(* Logix 5000 project; controller NWGG 1756-L72 rev 35.12; software revision 35.00; part 13 of 19 *)
(* tags used below, declared in another part *)
   tmrWeightTest : TIMER;
   Weight_Seed : DINT;
   _103_TANK_42_RECEIVING_LEG_RUNNING : BOOL;
   _106_TANK_17_AUGER_RUNNING : BOOL;
   _107_TANKS_1THRU7_SOUTH_RUNNING : BOOL;
   _108_CENTER_BELT_RUNNING : BOOL;
   _109_RAW_RECEIVING_NORTH_BELT_RUNNING : BOOL;
   _110_TANK_16_AUGER_RUNNING : BOOL;
   _113_HIGHROLLER_TANKS_11TO15_RUNNING : BOOL;
   _114_TANKS_1THRU7_NORTH_RUNNING : BOOL;
   _11_TANK_41_42_HIGHROLLER_RUNNING : BOOL;
   _123_CLEAN_LEG_RUNNING : BOOL;
   _1_CLEAN_SEED_UPPER_BELT_RUNNING : BOOL;
   _35_JUMP_LEG_RUNNING : BOOL;
   _3_LOWER_TANK_CONVAYOR_24TO26_RUNNING : BOOL;
   _43_SCREENINGS_LEG_RUNNING : BOOL;
   _4_LOWER_TANK_CONVAYOR_21TO23_RUNNING : BOOL;
   _5_LOWER_CROSS_BELT_RUNNING : BOOL;
   _701_TRUCK_REVERSING_BELT_RUNNING : BOOL;
   _703_TREATER_JUMP_BELT_RUNNING : BOOL;
   _9_TREATER_CONVAYOR_RUNNING : BOOL;
   Analog : AI[160];
   Calibration_Max : REAL;
   InEUMax : REAL;
   TestTag : REAL;
   Truck_Scales : udt_Truck_Scale[2];
(* MainProgram, continued *)

ROUTINE Totals   (* function block diagram *)
   SHEET 1
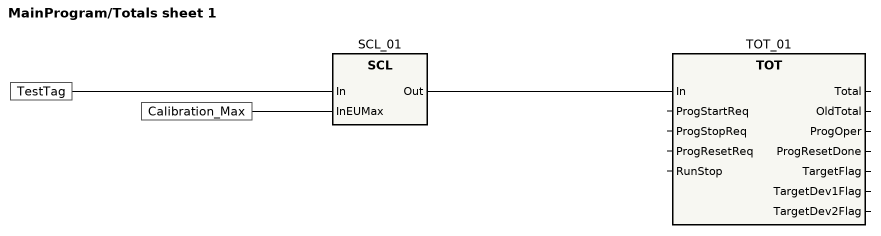
   SCL_01 : SCL(In := TestTag, InEUMax := Calibration_Max);
   TOT_01 : TOT(In := SCL_01.Out);   // unwired pins: ProgStartReq ProgStopReq ProgResetReq Total OldTotal ProgOper RunStop ProgResetDone TargetFlag TargetDev1Flag TargetDev2Flag
END_ROUTINE

ROUTINE VERIFACATION   (* ladder *)
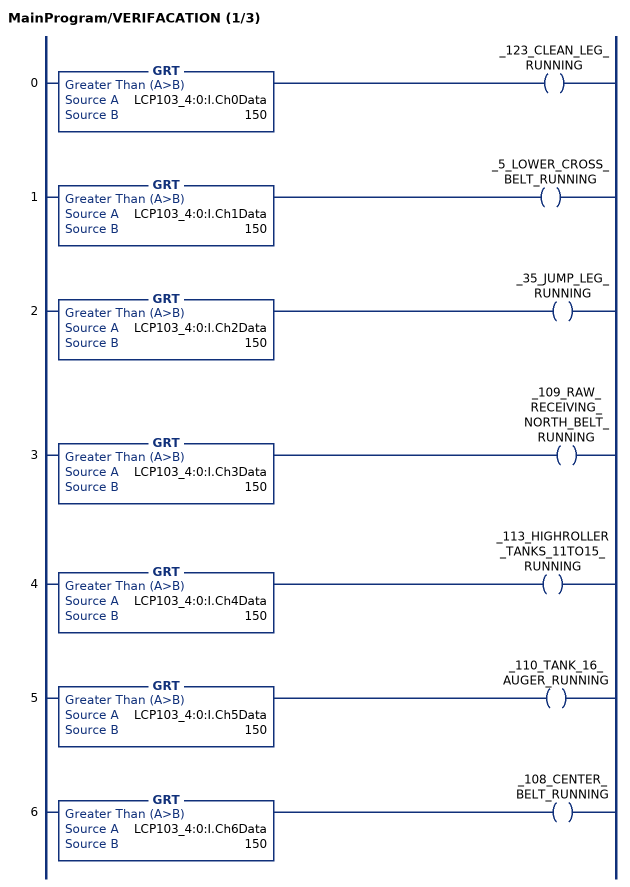
   0: GRT(LCP103_4:0:I.Ch0Data,150)OTE(_123_CLEAN_LEG_RUNNING);
   1: GRT(LCP103_4:0:I.Ch1Data,150)OTE(_5_LOWER_CROSS_BELT_RUNNING);
   2: GRT(LCP103_4:0:I.Ch2Data,150)OTE(_35_JUMP_LEG_RUNNING);
   3: GRT(LCP103_4:0:I.Ch3Data,150)OTE(_109_RAW_RECEIVING_NORTH_BELT_RUNNING);
   4: GRT(LCP103_4:0:I.Ch4Data,150)OTE(_113_HIGHROLLER_TANKS_11TO15_RUNNING);
   5: GRT(LCP103_4:0:I.Ch5Data,150)OTE(_110_TANK_16_AUGER_RUNNING);
   6: GRT(LCP103_4:0:I.Ch6Data,150)OTE(_108_CENTER_BELT_RUNNING);
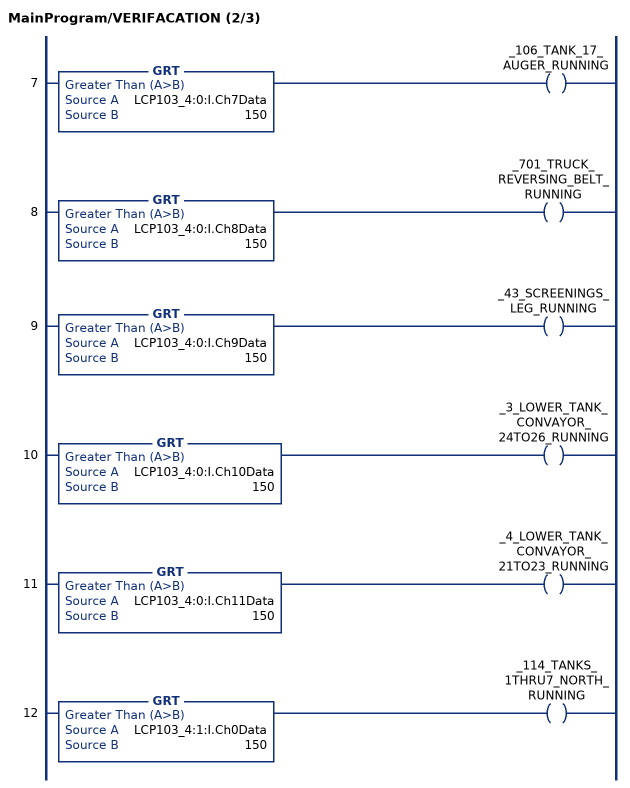
   7: GRT(LCP103_4:0:I.Ch7Data,150)OTE(_106_TANK_17_AUGER_RUNNING);
   8: GRT(LCP103_4:0:I.Ch8Data,150)OTE(_701_TRUCK_REVERSING_BELT_RUNNING);
   9: GRT(LCP103_4:0:I.Ch9Data,150)OTE(_43_SCREENINGS_LEG_RUNNING);
   10: GRT(LCP103_4:0:I.Ch10Data,150)OTE(_3_LOWER_TANK_CONVAYOR_24TO26_RUNNING);
   11: GRT(LCP103_4:0:I.Ch11Data,150)OTE(_4_LOWER_TANK_CONVAYOR_21TO23_RUNNING);
   12: GRT(LCP103_4:1:I.Ch0Data,150)OTE(_114_TANKS_1THRU7_NORTH_RUNNING);
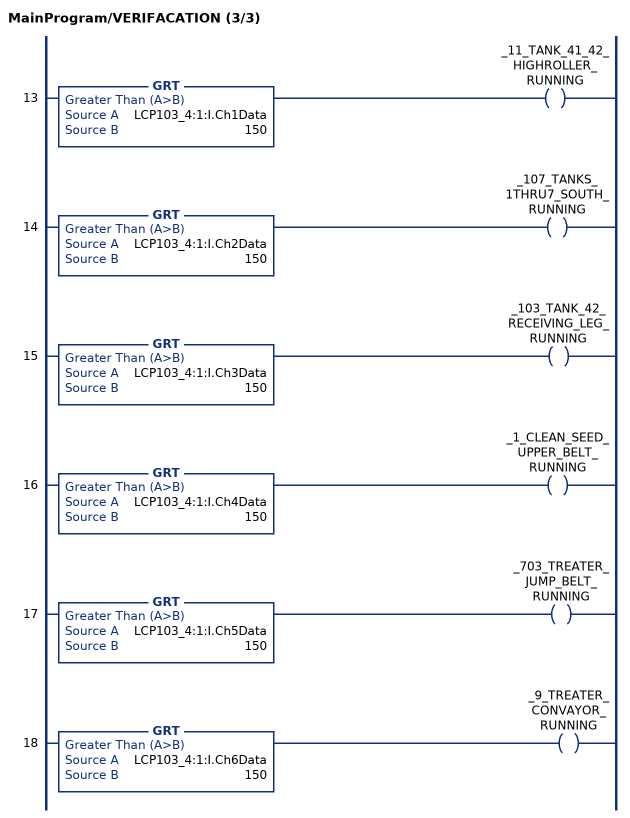
   13: GRT(LCP103_4:1:I.Ch1Data,150)OTE(_11_TANK_41_42_HIGHROLLER_RUNNING);
   14: GRT(LCP103_4:1:I.Ch2Data,150)OTE(_107_TANKS_1THRU7_SOUTH_RUNNING);
   15: GRT(LCP103_4:1:I.Ch3Data,150)OTE(_103_TANK_42_RECEIVING_LEG_RUNNING);
   16: GRT(LCP103_4:1:I.Ch4Data,150)OTE(_1_CLEAN_SEED_UPPER_BELT_RUNNING);
   17: GRT(LCP103_4:1:I.Ch5Data,150)OTE(_703_TREATER_JUMP_BELT_RUNNING);
   18: GRT(LCP103_4:1:I.Ch6Data,150)OTE(_9_TREATER_CONVAYOR_RUNNING);
END_ROUTINE

ROUTINE Weigh_Scales   (* ladder *)
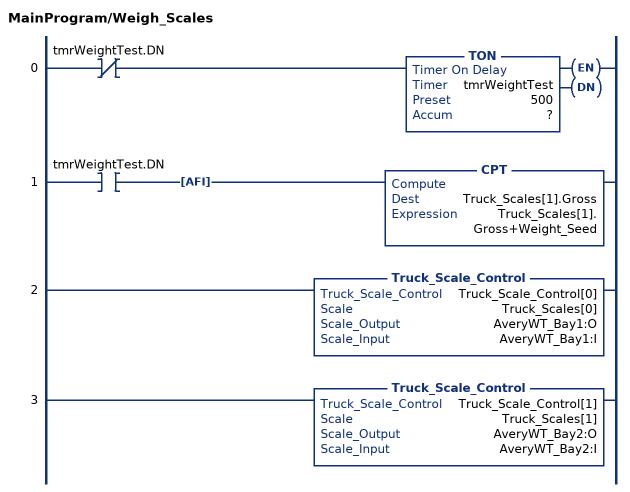
   0: XIO(tmrWeightTest.DN)TON(tmrWeightTest,?,?);
   1: XIC(tmrWeightTest.DN)AFI()CPT(Truck_Scales[1].Gross,Truck_Scales[1].Gross+Weight_Seed);
   2: Truck_Scale_Control(Truck_Scale_Control[0],Truck_Scales[0],AveryWT_Bay1:O,AveryWT_Bay1:I);
   3: Truck_Scale_Control(Truck_Scale_Control[1],Truck_Scales[1],AveryWT_Bay2:O,AveryWT_Bay2:I);
END_ROUTINE
END_PROGRAM

PROGRAM Scale   (* main routine MainRoutine *)
VAR
   ctlAddTime : CONTROL[2];
   ctrWtArray : COUNTER[2] := ([0].DN := 1, [1].DN := 1);
   Cur_Weight : REAL[2];
   Cur_Weight_Array_Idx : DINT := 16;
   Current_Gross : DINT[2];
   Current_Weight : REAL;
   Prev_Weight : REAL[2];
   Scale_Rate : REAL[2];
   Scale_Test_Rate_Mlt : DINT;
   ScaleIDX : DINT := 2;
   ShiftIDX : DINT := 20;
   TestRate : REAL[2];
   Time_Array : DINT[2,10] := ([0,0] := 9, [0,1] := 9, [0,2] := 10, [0,3] := 10, [0,4] := 8, [0,5] := 10, [0,6] := 9, [0,7] := 9, [0,8] := 9, [1,0] := 10, [1,1] := 9, [1,2] := 10, [1,3] := 10, [1,4] := 9, [1,5] := 10, [1,6] := 8, [1,7] := 10, [1,8] := 9);
   tmrRate : TIMER[2] := ([0].PRE := 1000, [0].ACC := 109, [0].EN := 1, [0].TT := 1, [1].PRE := 1000, [1].ACC := 126, [1].EN := 1, [1].TT := 1);
   tmrTestRate : TIMER[2] := ([1].ACC := 15, [1].EN := 1, [1].DN := 1);
   Total_Time : DINT[2];
   Weight_Array : REAL[2,40];
   Weight_Array_Idx : DINT[2] := ([0] := 14, [1] := 17);
   Weight_Array_Max : REAL[2];
   Weight_Sum : REAL[2];
END_VAR

ROUTINE AddWeights   (* ladder *)
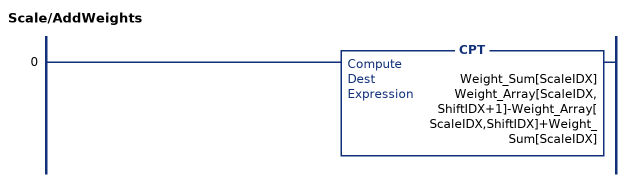
   0: CPT(Weight_Sum[ScaleIDX],Weight_Array[ScaleIDX,ShiftIDX+1]-Weight_Array[ScaleIDX,ShiftIDX]+Weight_Sum[ScaleIDX]);
END_ROUTINE

ROUTINE MainRoutine   (* ladder *)
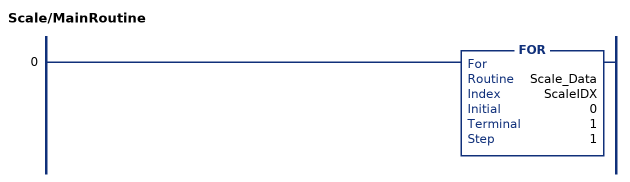
   0: FOR(Scale_Data,ScaleIDX,0,1,1);
END_ROUTINE

ROUTINE Scale_Data   (* ladder *)
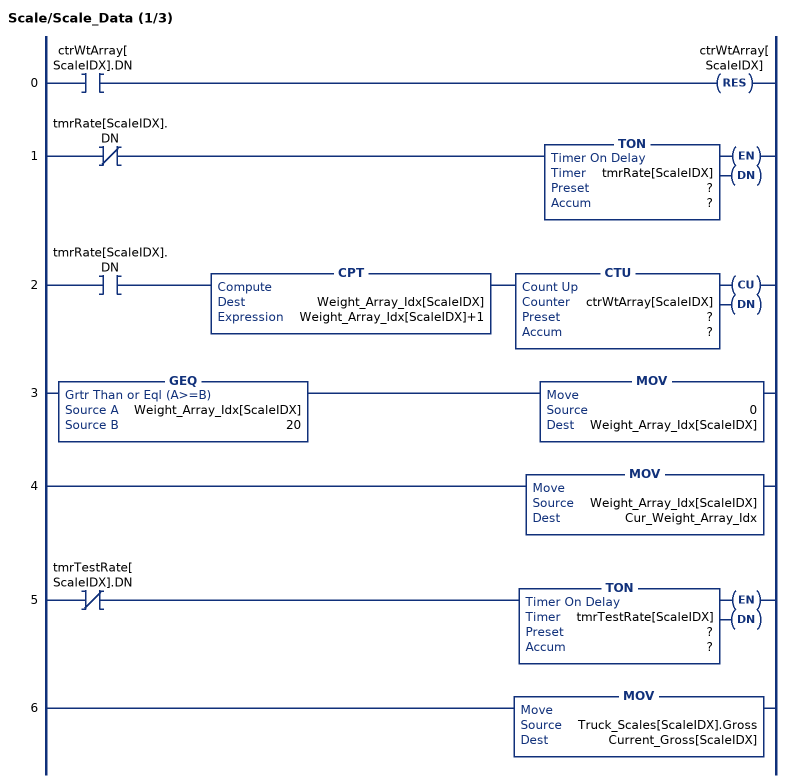
   0: XIC(ctrWtArray[ScaleIDX].DN)RES(ctrWtArray[ScaleIDX]);
   1: XIO(tmrRate[ScaleIDX].DN)TON(tmrRate[ScaleIDX],?,?);
   2: XIC(tmrRate[ScaleIDX].DN)CPT(Weight_Array_Idx[ScaleIDX],Weight_Array_Idx[ScaleIDX]+1)CTU(ctrWtArray[ScaleIDX],?,?);
   3: GEQ(Weight_Array_Idx[ScaleIDX],20)MOV(0,Weight_Array_Idx[ScaleIDX]);
   4: MOV(Weight_Array_Idx[ScaleIDX],Cur_Weight_Array_Idx);
   5: XIO(tmrTestRate[ScaleIDX].DN)TON(tmrTestRate[ScaleIDX],?,?);
   6: MOV(Truck_Scales[ScaleIDX].Gross,Current_Gross[ScaleIDX]);
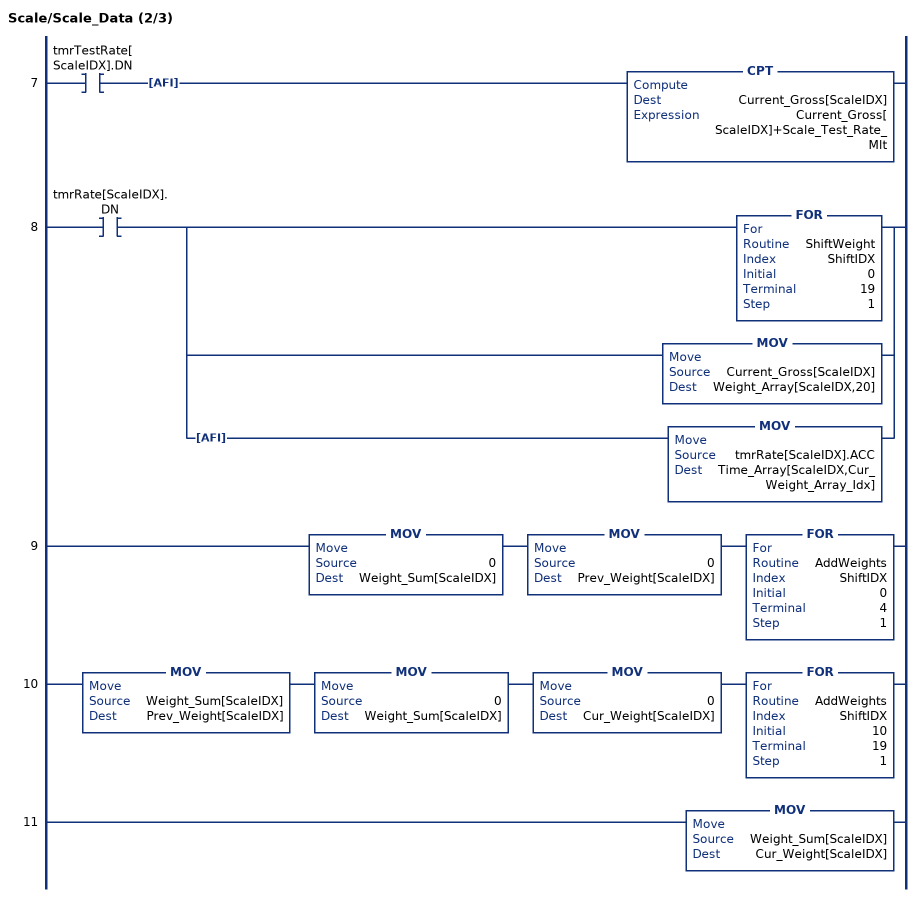
   7: XIC(tmrTestRate[ScaleIDX].DN)AFI()CPT(Current_Gross[ScaleIDX],Current_Gross[ScaleIDX]+Scale_Test_Rate_Mlt);
   8: XIC(tmrRate[ScaleIDX].DN)[FOR(ShiftWeight,ShiftIDX,0,19,1) ,MOV(Current_Gross[ScaleIDX],Weight_Array[ScaleIDX,20]) ,AFI() MOV(tmrRate[ScaleIDX].ACC,Time_Array[ScaleIDX,Cur_Weight_Array_Idx]) ];
   9: MOV(0,Weight_Sum[ScaleIDX])MOV(0,Prev_Weight[ScaleIDX])FOR(AddWeights,ShiftIDX,0,4,1);
   10: MOV(Weight_Sum[ScaleIDX],Prev_Weight[ScaleIDX])MOV(0,Weight_Sum[ScaleIDX])MOV(0,Cur_Weight[ScaleIDX])FOR(AddWeights,ShiftIDX,10,19,1);
   11: MOV(Weight_Sum[ScaleIDX],Cur_Weight[ScaleIDX]);
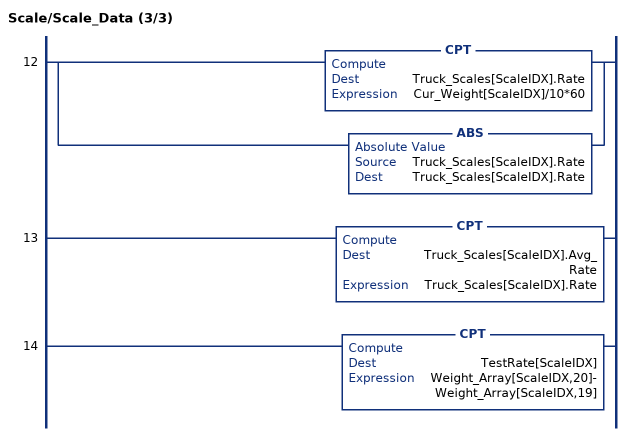
   12: [CPT(Truck_Scales[ScaleIDX].Rate,Cur_Weight[ScaleIDX]/10*60) ,ABS(Truck_Scales[ScaleIDX].Rate,Truck_Scales[ScaleIDX].Rate) ];
   13: CPT(Truck_Scales[ScaleIDX].Avg_Rate,Truck_Scales[ScaleIDX].Rate);
   14: CPT(TestRate[ScaleIDX],Weight_Array[ScaleIDX,20]-Weight_Array[ScaleIDX,19]);
END_ROUTINE

ROUTINE ShiftWeight   (* ladder *)
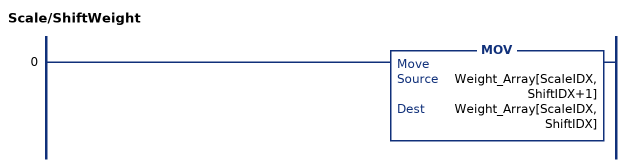
   0: MOV(Weight_Array[ScaleIDX,ShiftIDX+1],Weight_Array[ScaleIDX,ShiftIDX]);
END_ROUTINE
END_PROGRAM

PROGRAM SeedLoadoutMain   (* main routine MainRoutine *)
VAR
   Accept_Bin_Cal : BOOL;
   Air_Gates_Opened : BOOL;
   All_Stop : BOOL;
   ALM_Air_Gate_Failed_Open_Bin0 : ALARM_DIGITAL;
   ALM_Air_Gate_Failed_Open_Bin1 : ALARM_DIGITAL;
   ALM_Air_Gate_Failed_Open_Bin10 : ALARM_DIGITAL;
   ALM_Air_Gate_Failed_Open_Bin11 : ALARM_DIGITAL;
   ALM_Air_Gate_Failed_Open_Bin12 : ALARM_DIGITAL;
   ALM_Air_Gate_Failed_Open_Bin13 : ALARM_DIGITAL;
   ALM_Air_Gate_Failed_Open_Bin14 : ALARM_DIGITAL;
   ALM_Air_Gate_Failed_Open_Bin15 : ALARM_DIGITAL;
   ALM_Air_Gate_Failed_Open_Bin16 : ALARM_DIGITAL;
   ALM_Air_Gate_Failed_Open_Bin17 : ALARM_DIGITAL;
   ALM_Air_Gate_Failed_Open_Bin18 : ALARM_DIGITAL;
   ALM_Air_Gate_Failed_Open_Bin19 : ALARM_DIGITAL;
   ALM_Air_Gate_Failed_Open_Bin2 : ALARM_DIGITAL;
   ALM_Air_Gate_Failed_Open_Bin20 : ALARM_DIGITAL;
   ALM_Air_Gate_Failed_Open_Bin21 : ALARM_DIGITAL;
   ALM_Air_Gate_Failed_Open_Bin22 : ALARM_DIGITAL;
   ALM_Air_Gate_Failed_Open_Bin23 : ALARM_DIGITAL;
   ALM_Air_Gate_Failed_Open_Bin24 : ALARM_DIGITAL;
   ALM_Air_Gate_Failed_Open_Bin25 : ALARM_DIGITAL;
   ALM_Air_Gate_Failed_Open_Bin26 : ALARM_DIGITAL;
   ALM_Air_Gate_Failed_Open_Bin27 : ALARM_DIGITAL;
   ALM_Air_Gate_Failed_Open_Bin28 : ALARM_DIGITAL;
   ALM_Air_Gate_Failed_Open_Bin3 : ALARM_DIGITAL;
   ALM_Air_Gate_Failed_Open_Bin4 : ALARM_DIGITAL;
   ALM_Air_Gate_Failed_Open_Bin5 : ALARM_DIGITAL;
   ALM_Air_Gate_Failed_Open_Bin6 : ALARM_DIGITAL;
   ALM_Air_Gate_Failed_Open_Bin7 : ALARM_DIGITAL;
   ALM_Air_Gate_Failed_Open_Bin8 : ALARM_DIGITAL;
   ALM_Air_Gate_Failed_Open_Bin9 : ALARM_DIGITAL;
   ALM_K_Valve1_Treat_Failed : ALARM_DIGITAL;
   ALM_KValve0_Clean_Failed : ALARM_DIGITAL;
   ALM_KValve0_Treat_Failed : ALARM_DIGITAL;
   ALM_KValve1_Clean_Failed : ALARM_DIGITAL;
   ALM_NOT_USED : ALARM_DIGITAL;
   ALM_OVRAMP_Belt10 : ALARM_DIGITAL;
   ALM_OVRAMP_Belt11 : ALARM_DIGITAL;
   ALM_OVRAMP_Belt2 : ALARM_DIGITAL;
   ALM_OVRAMP_Belt3 : ALARM_DIGITAL;
   ALM_OVRAMP_Belt4 : ALARM_DIGITAL;
   ALM_OVRAMP_Belt5 : ALARM_DIGITAL;
   ALM_OVRAMP_Belt6 : ALARM_DIGITAL;
   ALM_OVRAMP_Belt7 : ALARM_DIGITAL;
   ALM_OVRAMP_Belt8 : ALARM_DIGITAL;
   ALM_OVRAMP_Belt9 : ALARM_DIGITAL;
   ALM_OVRAMP_CPLeg : ALARM_DIGITAL;
   ALM_PLUG_Belt1 : ALARM_DIGITAL;
   ALM_PLUG_Belt10 : ALARM_DIGITAL;
   ALM_PLUG_Belt11 : ALARM_DIGITAL;
   ALM_PLUG_Belt2 : ALARM_DIGITAL;
   ALM_PLUG_Belt3 : ALARM_DIGITAL;
   ALM_PLUG_Belt4 : ALARM_DIGITAL;
   ALM_PLUG_Belt5 : ALARM_DIGITAL;
   ALM_PLUG_Belt6 : ALARM_DIGITAL;
   ALM_PLUG_Belt7 : ALARM_DIGITAL;
   ALM_PLUG_Belt8 : ALARM_DIGITAL;
   ALM_PLUG_Belt9 : ALARM_DIGITAL;
   ALM_PLUG_CPLeg : ALARM_DIGITAL;
   ALM_SLP10_Belt1 : ALARM_DIGITAL;
   ALM_SLP10_Belt10 : ALARM_DIGITAL;
   ALM_SLP10_Belt11 : ALARM_DIGITAL;
   ALM_SLP10_Belt2 : ALARM_DIGITAL;
   ALM_SLP10_Belt3 : ALARM_DIGITAL;
   ALM_SLP10_Belt4 : ALARM_DIGITAL;
   ALM_SLP10_Belt5 : ALARM_DIGITAL;
   ALM_SLP10_Belt6 : ALARM_DIGITAL;
   ALM_SLP10_Belt7 : ALARM_DIGITAL;
   ALM_SLP10_Belt8 : ALARM_DIGITAL;
   ALM_SLP10_Belt9 : ALARM_DIGITAL;
   ALM_SLP10_CPLeg : ALARM_DIGITAL;
   ALM_SLP20_Belt1 : ALARM_DIGITAL;
   ALM_SLP20_Belt10 : ALARM_DIGITAL;
   ALM_SLP20_Belt11 : ALARM_DIGITAL;
   ALM_SLP20_Belt2 : ALARM_DIGITAL;
   ALM_SLP20_Belt3 : ALARM_DIGITAL;
   ALM_SLP20_Belt4 : ALARM_DIGITAL;
   ALM_SLP20_Belt5 : ALARM_DIGITAL;
   ALM_SLP20_Belt6 : ALARM_DIGITAL;
   ALM_SLP20_Belt7 : ALARM_DIGITAL;
   ALM_SLP20_Belt8 : ALARM_DIGITAL;
   ALM_SLP20_Belt9 : ALARM_DIGITAL;
   ALM_SLP20_CPLeg : ALARM_DIGITAL;
   ALM_WONT_START_Belt1 : ALARM_DIGITAL;
   ALM_WONT_START_Belt10 : ALARM_DIGITAL;
   ALM_WONT_START_Belt11 : ALARM_DIGITAL;
   ALM_WONT_START_Belt2 : ALARM_DIGITAL;
   ALM_WONT_START_Belt3 : ALARM_DIGITAL;
   ALM_WONT_START_Belt4 : ALARM_DIGITAL;
   ALM_WONT_START_Belt5 : ALARM_DIGITAL;
   ALM_WONT_START_Belt6 : ALARM_DIGITAL;
   ALM_WONT_START_Belt7 : ALARM_DIGITAL;
   ALM_WONT_START_Belt8 : ALARM_DIGITAL;
   ALM_WONT_START_Belt9 : ALARM_DIGITAL;
   ALM_WONT_START_CPLeg : ALARM_DIGITAL;
   Always_Off : BOOL;
   Andco_Auto_Mode : BOOL;
   Andco_Rate : DINT;
   Auto_Mode : BOOL := 1;
   Auto_Mode_ONS : BOOL;
   Auto_Start_Reversing_Belt_Fans : BOOL;
   Auto_Start_Treatment : BOOL;
   Auto_Stop_Clean : BOOL;
   Auto_Stop_Clean_Belt_11 : BOOL;
   Auto_Stop_Transfer : BOOL;
   Auto_Stop_Treat : BOOL;
   Available_For_Clean_Loadout : DINT := 536870911;
   Available_For_Treat_Loadout : DINT := 536870911;
   b3 : ALARM_DIGITAL;
   B_Offset : REAL;
   Batch_Status : DINT;
   BC_3_Belt_Required : BOOL;
   BC_9_Interlock : BOOL;
   Belt : udt_Motor[16] := ([0].Motor_Start.Auto_Stop_Delay := 5000, [1].Motor_Start.Auto_Stop_Delay := 5000, [1].Motor_Control.Spd_10_Pct := 1, [1].Motor_Control.Motor_Amps := -0.32500002, [1].Motor_Control.Motor_Batch_Ready := 1, [1].Motor_Control.Motor_Batch_Ready_Clean := 1, [1].Motor_Control.Motor_Batch_Ready_Treat := 1, [1].Motor_Control.Motor_Batch_Ready_Transfer := 1, [1].Motor_Config.Definition := 'Middle Concrete', [1].Motor_Config.Wind_Up_Time := 3000, [1].Motor_Config.Stop_At_SLP20 := 1, [1].Motor_Config.Stop_At_Max_Amps := 1, [1].Motor_Config.Max_Amps := 1000.0, [2].Motor_Start.Auto_Stop_Delay := 5000, [2].Motor_Control.Spd_10_Pct := 1, [2].Motor_Control.Motor_Amps := -0.4125, [2].Motor_Control.Motor_Batch_Ready := 1, [2].Motor_Control.Motor_Batch_Ready_Clean := 1, [2].Motor_Control.Motor_Batch_Ready_Treat := 1, [2].Motor_Control.Motor_Batch_Ready_Transfer := 1, [2].Motor_Config.Definition := 'North Concrete', [2].Motor_Config.Wind_Up_Time := 3000, [2].Motor_Config.Stop_At_SLP20 := 1, [3].Motor_Start.Auto_Stop_Delay := 5000, [3].Motor_Control.Spd_10_Pct := 1, [3].Motor_Control.Motor_Amps := -0.5125, [3].Motor_Control.Motor_Batch_Ready := 1, [3].Motor_Control.Motor_Batch_Ready_Clean := 1, [3].Motor_Control.Motor_Batch_Ready_Treat := 1, [3].Motor_Control.Motor_Batch_Ready_Transfer := 1, [3].Motor_Config.Definition := 'South Concrete', [3].Motor_Config.Wind_Up_Time := 3000, [3].Motor_Config.Stop_At_SLP20 := 1, [4].Motor_Start.Auto_Stop_Delay := 5000, [4].Motor_Control.Motor_Amps := -0.05285539, [4].Motor_Control.Motor_Batch_Ready := 1, [4].Motor_Control.Motor_Batch_Ready_Clean := 1, [4].Motor_Control.Motor_Batch_Ready_Treat := 1, [4].Motor_Control.Motor_Batch_Ready_Transfer := 1, [4].Motor_Config.Definition := 'Reversing', [4].Motor_Config.Wind_Up_Time := 6000, [4].Motor_Config.Stop_At_SLP20 := 1, [5].Motor_Start.Auto_Stop_Delay := 5000, [5].Motor_Control.Spd_10_Pct := 1, [5].Motor_Control.Motor_Amps := 0.018231237, [5].Motor_Control.Motor_Batch_Ready := 1, [5].Motor_Control.Motor_Batch_Ready_Clean := 1, [5].Motor_Control.Motor_Batch_Ready_Treat := 1, [5].Motor_Control.Motor_Batch_Ready_Transfer := 1, [5].Motor_Config.Definition := 'Treat Jump', [5].Motor_Config.Wind_Up_Time := 3000, [5].Motor_Config.Stop_At_SLP20 := 1, [6].Motor_Start.Auto_Stop_Delay := 5000, [6].Motor_Control.Spd_10_Pct := 1, [6].Motor_Control.Motor_Amps := 0.013243717, [6].Motor_Control.Motor_Batch_Ready := 1, [6].Motor_Control.Motor_Batch_Ready_Clean := 1, [6].Motor_Control.Motor_Batch_Ready_Treat := 1, [6].Motor_Control.Motor_Batch_Ready_Transfer := 1, [6].Motor_Config.Definition := 'Clean Jump',
        [6].Motor_Config.Wind_Up_Time := 3000, [6].Motor_Config.Stop_At_SLP20 := 1, [6].Motor_Config.Plugged_Sensor_Disabled := 1, [7].Motor_Start.Auto_Stop_Delay := 5000, [7].Motor_Control.Spd_10_Pct := 1, [7].Motor_Control.Motor_Amps := -0.23403546, [7].Motor_Control.Motor_Batch_Ready := 1, [7].Motor_Control.Motor_Batch_Ready_Clean := 1, [7].Motor_Control.Motor_Batch_Ready_Treat := 1, [7].Motor_Control.Motor_Batch_Ready_Transfer := 1, [7].Motor_Config.Definition := 'BC-9', [7].Motor_Config.Wind_Up_Time := 3000, [7].Motor_Config.Stop_At_SLP20 := 1, [7].Motor_Config.Plugged_Sensor_Disabled := 1, [8].Motor_Start.Auto_Stop_Delay := 5000, [8].Motor_Control.Spd_20_Pct := 1, [8].Motor_Control.Motor_Amps := 0.001667556, [8].Motor_Control.Motor_Batch_Ready := 1, [8].Motor_Control.Motor_Batch_Ready_Clean := 1, [8].Motor_Control.Motor_Batch_Ready_Treat := 1, [8].Motor_Control.Motor_Batch_Ready_Transfer := 1, [8].Motor_Config.Definition := 'BC-4', [8].Motor_Config.Wind_Up_Time := 3000, [8].Motor_Config.Speed_Sensor_Disabled := 1, [8].Motor_Config.Plugged_Sensor_Disabled := 1, [9].Motor_Start.Auto_Stop_Delay := 5000, [9].Motor_Control.Spd_20_Pct := 1, [9].Motor_Control.Motor_Amps := 0.033333335, [9].Motor_Control.Motor_Batch_Ready := 1, [9].Motor_Control.Motor_Batch_Ready_Clean := 1, [9].Motor_Control.Motor_Batch_Ready_Treat := 1, [9].Motor_Control.Motor_Batch_Ready_Transfer := 1, [9].Motor_Config.Definition := 'BC-3', [9].Motor_Config.Wind_Up_Time := 3000, [10].Motor_Start.Auto_Stop_Delay := 5000, [10].Motor_Control.Spd_20_Pct := 1, [10].Motor_Control.Motor_Amps := 0.016583197, [10].Motor_Control.Motor_Batch_Ready := 1, [10].Motor_Control.Motor_Batch_Ready_Clean := 1, [10].Motor_Control.Motor_Batch_Ready_Treat := 1, [10].Motor_Control.Motor_Batch_Ready_Transfer := 1, [10].Motor_Config.Definition := 'High Roller', [10].Motor_Config.Wind_Up_Time := 3000, [11].Motor_Start.Auto_Stop_Delay := 5000, [11].Motor_Control.Spd_20_Pct := 1, [11].Motor_Control.Motor_Amps := -0.008290774, [11].Motor_Control.Motor_Batch_Ready := 1, [11].Motor_Control.Motor_Batch_Ready_Clean := 1, [11].Motor_Control.Motor_Batch_Ready_Treat := 1, [11].Motor_Control.Motor_Batch_Ready_Transfer := 1, [11].Motor_Config.Definition := 'BC-5', [11].Motor_Config.Wind_Up_Time := 3000, [12].Motor_Start.Auto_Stop_Delay := 5000);
   Belt_Amps_Scale : SCALE[11];
   Belt_Gate_Leg_ON : BOOL;
   Belts_Ready : BOOL := 1;
   Belts_Running : BOOL;
   Bin_Cal : BOOL;
   Bin_Cal_IDX : DINT := -1;
   Bin_Calibration : BOOL;
   Bin_Clean_Pause : BOOL;
   Bin_Gate_Test : BOOL := 1;
   Bin_Loadout_Control : Loadout_Bin_Control[29] := ([0].Use_Bindicator := 1, [0].RawAnalogTag := 10270, [1].RawAnalogTag := 9993, [2].Use_Bindicator := 1, [2].RawAnalogTag := 8109, [3].RawAnalogTag := 3610, [4].RawAnalogTag := 7694, [5].RawAnalogTag := 5041, [6].RawAnalogTag := 9661, [7].RawAnalogTag := 9884, [8].RawAnalogTag := 10717, [9].RawAnalogTag := 9078, [10].RawAnalogTag := 8853, [11].RawAnalogTag := 9587, [12].RawAnalogTag := 7657, [13].RawAnalogTag := 9087, [14].RawAnalogTag := 9078, [15].RawAnalogTag := 8853, [16].Use_Bindicator := 1, [16].RawAnalogTag := 14748, [17].Use_Bindicator := 1, [17].RawAnalogTag := 15440, [18].Use_Bindicator := 1, [18].RawAnalogTag := 14244, [19].Use_Bindicator := 1, [19].RawAnalogTag := 13454, [20].Use_Bindicator := 1, [20].RawAnalogTag := 14460, [21].Use_Auger_Relay := 1, [21].Use_Bindicator := 1, [21].RawAnalogTag := 6343, [22].Use_Auger_Relay := 1, [22].Use_Bindicator := 1, [22].RawAnalogTag := 8758, [23].Use_Bindicator := 1, [23].RawAnalogTag := 15944, [24].Use_Bindicator := 1, [24].RawAnalogTag := 15184, [25].Use_Bindicator := 1, [25].RawAnalogTag := 15745, [26].Use_Bindicator := 1, [26].RawAnalogTag := 15279, [27].Use_Bindicator := 1, [27].RawAnalogTag := 14611, [28].Use_Bindicator := 1, [28].RawAnalogTag := 15145);
   Bin_Open_test : BOOL := 1;
   Bin_Transfer_Pause : BOOL;
   Bin_Treat_Pause : BOOL;
   Bin_Use_Index : DINT;
   Bin_Variety_Id : STRING[30] := ([0] := '823048', [1] := '823054', [2] := '823058', [3] := '823038', [4] := '823082', [5] := '823090', [6] := '823054', [7] := '823001', [9] := '873002', [10] := '873002', [11] := '873003', [12] := '823072', [16] := '823098', [17] := '843022', [19] := '822087', [20] := '803003', [21] := '823093', [22] := '843036', [23] := '843001', [24] := '843002', [25] := '843022', [26] := '803003', [27] := '823087', [28] := '803021');
   Bins_Rqd : BOOL;
   Blow_Out_Time : DINT;
   Blow_Out_Time_Remaining : REAL := -0.016;
   Blower_707_Running : BOOL;
   boolTransferTime : BOOL;
   Cal_Bin_Status : DINT;
   Cal_Done : BOOL;
   Calibrate_Mode : BOOL;
   Cancel_Bin_Config : BOOL;
   ckIDX : DINT := 29;
   Clean_Batch_Status : DINT;
   Clean_Bin_Gates_Opened : BOOL := 1;
   Clean_Interlock : BOOL;
   Clean_K_Relay_Not_Used : BOOL := 1;
   Clean_Load_Requested : BOOL;
   Clean_Scale_Target : DINT;
   Clean_Scale_Unavailable : BOOL;
   CleanHours : DINT;
   CleanMinuets : DINT;
   CleanSeconds : DINT;
   cntCleanTime : COUNTER := (PRE := 1);
   cntTest : COUNTER := (PRE := 100, ACC := 4);
   cntTransferTime : COUNTER := (PRE := 1);
   cntTreatTime : COUNTER := (PRE := 1);
   Concrete_Belts_Ready : BOOL;
   Concrete_Bin_Timing_Offset : DINT := 5;
   Concrete_Clean_Belts_Ready : BOOL;
   Concrete_Fan_Start : BOOL;
   Concrete_Leg : udt_Motor := (Motor_Start.Auto_Stop_Delay := 1, Motor_Control.Spd_20_Pct := 1, Motor_Control.Spd_10_Pct := 1, Motor_Control.Motor_Amps := -0.4625, Motor_Control.Motor_Batch_Ready_Clean := 1, Motor_Control.Motor_Batch_Ready_Treat := 1, Motor_Control.Motor_Batch_Ready_Transfer := 1, Motor_Config.Definition := 'CONCRETE LEG', Motor_Config.Wind_Up_Time := 4000, Motor_Config.Speed_Sensor_Disabled := 1, Motor_Config.Plugged_Sensor_Disabled := 1);
   Concrete_Leg_Interlock : BOOL;
   Concrete_Leg_Rqd : BOOL;
   Config_Bin_Name : STRING;
   Config_Cancel_Bin : BOOL := 1;
   Config_Class : STRING;
   Config_Clean_Delay_Start : REAL;
   Config_Clean_Delay_Stop : REAL;
   Config_Item_Number : STRING;
   Config_Name : STRING;
   Config_Pounds_Per_Inch : REAL;
   Config_Save_Bin : BOOL;
   Config_Treat_Delay_Start : REAL;
   Config_Treat_Delay_Stop : REAL;
   Configure_Clean_Delay : DINT := 36000;
   Configure_LoadoutBin : udt_Loadout_Bin := (Bin_Description := '9', Bin_Variety.Item_Number := '382010', Clean_Load_Delay_Start := 36000, Treat_Load_Delay_Start := 36000, Andco_Values.Raw_Position := 7, Andco_Values.Max_Position := 103, Andco_Values.Preact := 3, Andco_Values.Percent_Open := 0.067961164, Andco_Values.New_Pos := 9, Andco_Values.Width := 6.0);
   Configure_Treat_Delay_Start : DINT := 36000;
   ConfigureIndex : DINT := -1;
   ConfirmStop : BOOL;
   Current_Dist_List_IDX : DINT := 15;
   Current_Dist_Position : STRING := '10';
   Current_Longest_Time : DINT;
   Current_System_Msg_idx : DINT;
   Current_Transfer_Bin_From : BOOL[32];
   Current_Transfer_Bin_To : BOOL[32];
   DeltaX : REAL := -3028.0;
   DeltaY : REAL := -1000.0;
   Empty_String : STRING; {constant}
   Empty_Variety_ID : STRING := '0'; {constant}
   Finish_Treat_Ok : BOOL;
   FSC_Reverse : CONTROL;
   High_Roller_Belt_Bins_Required : BOOL;
   IDX : DINT := 29;
   Interlock_Not_Used : BOOL := 1;
   loa : ALARM_DIGITAL;
   Loadout_Bin : udt_Loadout_Bin[29] := ([0].Bin_Description := '3', [0].Bin_Variety.Item_Number := '823048', [0].Bin_Variety.Name := 'SEAHAWK CERTIFIED SPRING SWH', [0].Bin_Variety.Class := 'Certified', [0].Rate_Cal_Points[1].Andco_Position := 3631, [0].Rate_Cal_Points[1].Rate := 1000, [0].Rate_Cal_Points[2].Andco_Position := 6242, [0].Rate_Cal_Points[2].Rate := 2000, [0].Rate_Cal_Points[3].Andco_Position := 7451, [0].Rate_Cal_Points[3].Rate := 3000, [0].Rate_Cal_Points[4].Andco_Position := 9390, [0].Rate_Cal_Points[4].Rate := 4000, [0].Clean_Load_Delay_Start := 36050, [0].Treat_Load_Delay_Start := 29000, [0].Andco_Values.Cal_Status := 4, [0].Andco_Values.Raw_Position := 9707, [0].Andco_Values.Max_Position := 15761, [0].Andco_Values.Preact := 20, [0].Andco_Values.Percent_Open := 0.63870245, [0].Andco_Values.New_Pos := 1, [0].Andco_Values.Width := 6.0, [0].Andco_Values.Rate := 4163.4863, [0].Andco_Values.Pounds_Per_Inch := 65.0, [0].Andco_Values.New_Rate := 20.0, [0].Andco_Values.Analog := 1, [0].Andco_Values.Min_Position := 563, [0].Andco_Values.Length := 12.0, [0].Andco_Values.InchesOpen := 7.6644297, [0].Andco_Values.AnalogValue := 10270, [0].Clean_Load_Delay_Stop := 36050, [0].Treat_Load_Delay_Stop := 32000, [0].tmrStopDelay.EN := 1, [0].tmrStopDelay.TT := 1, [0].Available_For_Clean_Load := 1, [0].Available_For_Treat_Load := 1, [1].Bin_Description := '1', [1].Bin_Variety.Item_Number := '823054', [1].Bin_Variety.Name := 'RYAN CERTIFIED SPRING SWH', [1].Bin_Variety.Class := 'Certified', [1].Bin_Variety.Color[0].Color := 1, [1].Rate_Cal_Points[1].Andco_Position := 3454, [1].Rate_Cal_Points[1].Rate := 1000, [1].Rate_Cal_Points[2].Andco_Position := 5979, [1].Rate_Cal_Points[2].Rate := 2000, [1].Rate_Cal_Points[3].Andco_Position := 7870, [1].Rate_Cal_Points[3].Rate := 3000, [1].Rate_Cal_Points[4].Andco_Position := 9015, [1].Rate_Cal_Points[4].Rate := 4000, [1].Clean_Load_Delay_Start := 36100, [1].Treat_Load_Delay_Start := 29000, [1].Andco_Values.Cal_Status := 2, [1].Andco_Values.Raw_Position := 9424, [1].Andco_Values.Max_Position := 14962, [1].Andco_Values.Preact := 20, [1].Andco_Values.Percent_Open := 0.65476274, [1].Andco_Values.New_Pos := 2, [1].Andco_Values.Width := 6.0, [1].Andco_Values.Rate := 4357.205, [1].Andco_Values.Pounds_Per_Inch := 86.6, [1].Andco_Values.New_Rate := 1.0,
        [1].Andco_Values.Analog := 1, [1].Andco_Values.Min_Position := 569, [1].Andco_Values.Length := 12.0, [1].Andco_Values.InchesOpen := 7.857153, [1].Andco_Values.AnalogValue := 9993, [1].Clean_Load_Delay_Stop := 35000, [1].Treat_Load_Delay_Stop := 35000, [1].tmrStartDelay.PRE := 3000, [1].tmrStopDelay.PRE := 1000, [1].tmrStopDelay.EN := 1, [1].tmrStopDelay.TT := 1, [1].StartDelayPre := 3000, [1].StopDelayPre := 1000, [1].Available_For_Clean_Load := 1, [1].Available_For_Treat_Load := 1, [2].Bin_Description := '11', [2].Bin_Variety.Item_Number := '823058', [2].Bin_Variety.Name := 'MPRESS CERTIFIED FALL SWH', [2].Bin_Variety.Class := 'Certified', [2].Bin_Variety.Color[0].Color := 1, [2].Rate_Cal_Points[1].Andco_Position := 3384, [2].Rate_Cal_Points[1].Rate := 1000, [2].Rate_Cal_Points[2].Andco_Position := 5322, [2].Rate_Cal_Points[2].Rate := 2000, [2].Rate_Cal_Points[3].Andco_Position := 6882, [2].Rate_Cal_Points[3].Rate := 3000, [2].Rate_Cal_Points[4].Andco_Position := 7544, [2].Rate_Cal_Points[4].Rate := 4000, [2].Clean_Load_Delay_Start := 36000, [2].Treat_Load_Delay_Start := 30000, [2].Andco_Values.Cal_Status := 2, [2].Andco_Values.Raw_Position := 7352, [2].Andco_Values.Max_Position := 13688, [2].Andco_Values.Preact := 20, [2].Andco_Values.Percent_Open := 0.5686002, [2].Andco_Values.New_Pos := 54, [2].Andco_Values.Width := 6.0, [2].Andco_Values.Rate := 3709.9697, [2].Andco_Values.Pounds_Per_Inch := 65.0, [2].Andco_Values.New_Rate := 4000.0, [2].Andco_Values.Analog := 1, [2].Andco_Values.Min_Position := 758, [2].Andco_Values.Length := 12.0, [2].Andco_Values.InchesOpen := 6.823202, [2].Andco_Values.AnalogValue := 8110, [2].Clean_Load_Delay_Stop := 36000, [2].Treat_Load_Delay_Stop := 33000, [2].tmrStopDelay.EN := 1, [2].tmrStopDelay.TT := 1, [2].Available_For_Clean_Load := 1, [2].Available_For_Treat_Load := 1, [3].Bin_Description := '9', [3].Bin_Variety.Item_Number := '823038', [3].Bin_Variety.Name := 'DRIVE CERTIFIED FALL SWH', [3].Bin_Variety.Class := 'Certified', [3].Bin_Variety.Color[0].Color := 1, [3].Rate_Cal_Points[1].Andco_Position := 1926, [3].Rate_Cal_Points[1].Rate := 1000, [3].Rate_Cal_Points[2].Andco_Position := 5008, [3].Rate_Cal_Points[2].Rate := 2000,
        [3].Rate_Cal_Points[3].Andco_Position := 6109, [3].Rate_Cal_Points[3].Rate := 3000, [3].Rate_Cal_Points[4].Andco_Position := 7052, [3].Rate_Cal_Points[4].Rate := 4000, [3].Clean_Load_Delay_Start := 36000, [3].Treat_Load_Delay_Start := 31000, [3].Andco_Values.Cal_Status := 2, [3].Andco_Values.Raw_Position := 3192, [3].Andco_Values.Max_Position := 13763, [3].Andco_Values.Preact := 20, [3].Andco_Values.Percent_Open := 0.23919071, [3].Andco_Values.Width := 6.0, [3].Andco_Values.Rate := 1410.7722, [3].Andco_Values.Pounds_Per_Inch := 65.0, [3].Andco_Values.Analog := 1, [3].Andco_Values.Min_Position := 418, [3].Andco_Values.Length := 12.0, [3].Andco_Values.InchesOpen := 2.8702886, [3].Andco_Values.AnalogValue := 3610, [3].Clean_Load_Delay_Stop := 36000, [3].Treat_Load_Delay_Stop := 34000, [3].tmrStopDelay.EN := 1, [3].tmrStopDelay.TT := 1, [3].Available_For_Clean_Load := 1, [3].Available_For_Treat_Load := 1, [4].Bin_Description := '5', [4].Bin_Variety.Item_Number := '823082', [4].Bin_Variety.Name := 'LCS DAGGER AX - 5235 COAXIUM CERTIFIED SWH', [4].Bin_Variety.Class := 'Certified', [4].Rate_Cal_Points[1].Andco_Position := 3130, [4].Rate_Cal_Points[1].Rate := 1000, [4].Rate_Cal_Points[2].Andco_Position := 5282, [4].Rate_Cal_Points[2].Rate := 2000, [4].Rate_Cal_Points[3].Andco_Position := 6505, [4].Rate_Cal_Points[3].Rate := 3000, [4].Rate_Cal_Points[4].Andco_Position := 7576, [4].Rate_Cal_Points[4].Rate := 4000, [4].Clean_Load_Delay_Start := 36000, [4].Treat_Load_Delay_Start := 30000, [4].Andco_Values.Cal_Status := 4, [4].Andco_Values.Raw_Position := 7436, [4].Andco_Values.Max_Position := 13094, [4].Andco_Values.Preact := 20, [4].Andco_Values.Tolerance := 1, [4].Andco_Values.Percent_Open := 0.5793082, [4].Andco_Values.New_Pos := 63, [4].Andco_Values.Width := 6.0, [4].Andco_Values.Rate := 3869.281, [4].Andco_Values.Pounds_Per_Inch := 65.0, [4].Andco_Values.New_Rate := 4000.0, [4].Andco_Values.Analog := 1, [4].Andco_Values.Min_Position := 258, [4].Andco_Values.Length := 12.0, [4].Andco_Values.InchesOpen := 6.9516983, [4].Andco_Values.AnalogValue := 7694, [4].Clean_Load_Delay_Stop := 36000, [4].Treat_Load_Delay_Stop := 33000, [4].tmrStopDelay.EN := 1, [4].tmrStopDelay.TT := 1, [4].Available_For_Clean_Load := 1,
        [4].Available_For_Treat_Load := 1, [5].Bin_Description := '4', [5].Bin_Variety.Item_Number := '823090', [5].Bin_Variety.Name := 'REAPER-0293 CERTIFIED SWH', [5].Bin_Variety.Class := 'Certified', [5].Bin_Variety.Color[0].Color := 1, [5].Rate_Cal_Points[1].Andco_Position := 2925, [5].Rate_Cal_Points[1].Rate := 1000, [5].Rate_Cal_Points[2].Andco_Position := 4802, [5].Rate_Cal_Points[2].Rate := 2000, [5].Rate_Cal_Points[3].Andco_Position := 6340, [5].Rate_Cal_Points[3].Rate := 3000, [5].Rate_Cal_Points[4].Andco_Position := 7786, [5].Rate_Cal_Points[4].Rate := 4000, [5].Clean_Load_Delay_Start := 38000, [5].Treat_Load_Delay_Start := 30000, [5].Andco_Values.Cal_Status := 4, [5].Andco_Values.Raw_Position := 4496, [5].Andco_Values.Max_Position := 12868, [5].Andco_Values.Preact := 20, [5].Andco_Values.Percent_Open := 0.36484623, [5].Andco_Values.Width := 6.0, [5].Andco_Values.Rate := 1836.9739, [5].Andco_Values.Pounds_Per_Inch := 65.0, [5].Andco_Values.Analog := 1, [5].Andco_Values.Min_Position := 545, [5].Andco_Values.Length := 12.0, [5].Andco_Values.InchesOpen := 4.3781548, [5].Andco_Values.AnalogValue := 5041, [5].Clean_Load_Delay_Stop := 60000, [5].Treat_Load_Delay_Stop := 34000, [5].tmrStartDelay.PRE := 1000, [5].tmrStopDelay.EN := 1, [5].tmrStopDelay.TT := 1, [5].StartDelayPre := 1000, [5].Available_For_Clean_Load := 1, [5].Available_For_Treat_Load := 1, [6].Bin_Description := '7', [6].Bin_Variety.Item_Number := '823054', [6].Bin_Variety.Name := 'RYAN CERTIFIED SPRING SWH', [6].Bin_Variety.Class := 'Certified', [6].Bin_Variety.Color[0].Color := 1, [6].Rate_Cal_Points[1].Andco_Position := 3297, [6].Rate_Cal_Points[1].Rate := 1000, [6].Rate_Cal_Points[2].Andco_Position := 5415, [6].Rate_Cal_Points[2].Rate := 2000, [6].Rate_Cal_Points[3].Andco_Position := 7178, [6].Rate_Cal_Points[3].Rate := 3000, [6].Rate_Cal_Points[4].Andco_Position := 9109, [6].Rate_Cal_Points[4].Rate := 4000, [6].Clean_Load_Delay_Start := 36000, [6].Treat_Load_Delay_Start := 30000, [6].Andco_Values.Cal_Status := 4, [6].Andco_Values.Raw_Position := 9035, [6].Andco_Values.Max_Position := 15835, [6].Andco_Values.Preact := 20, [6].Andco_Values.Percent_Open := 0.5940171, [6].Andco_Values.New_Pos := 67, [6].Andco_Values.Width := 6.0, [6].Andco_Values.Rate := 3961.6777,
        [6].Andco_Values.Pounds_Per_Inch := 65.0, [6].Andco_Values.New_Rate := 4000.0, [6].Andco_Values.Analog := 1, [6].Andco_Values.Min_Position := 625, [6].Andco_Values.Length := 12.0, [6].Andco_Values.InchesOpen := 7.1282053, [6].Andco_Values.AnalogValue := 9660, [6].Clean_Load_Delay_Stop := 36000, [6].Treat_Load_Delay_Stop := 34000, [6].tmrStopDelay.EN := 1, [6].tmrStopDelay.TT := 1, [6].Available_For_Clean_Load := 1, [6].Available_For_Treat_Load := 1, [7].Bin_Description := '10', [7].Bin_Variety.Item_Number := '823001', [7].Bin_Variety.Name := 'ARTDECO CERTIFIED FALL SWH', [7].Bin_Variety.Class := 'Certified', [7].Bin_Variety.Color[0].Color := 1, [7].Rate_Cal_Points[1].Andco_Position := 3007, [7].Rate_Cal_Points[1].Rate := 1000, [7].Rate_Cal_Points[2].Andco_Position := 5443, [7].Rate_Cal_Points[2].Rate := 2000, [7].Rate_Cal_Points[3].Andco_Position := 7342, [7].Rate_Cal_Points[3].Rate := 3000, [7].Rate_Cal_Points[4].Andco_Position := 9304, [7].Rate_Cal_Points[4].Rate := 4000, [7].Clean_Load_Delay_Start := 36500, [7].Treat_Load_Delay_Start := 30000, [7].Andco_Values.Cal_Status := 4, [7].Andco_Values.Raw_Position := 9878, [7].Andco_Values.Max_Position := 10246, [7].Andco_Values.Preact := 20, [7].Andco_Values.Percent_Open := 0.9646484, [7].Andco_Values.New_Pos := 68, [7].Andco_Values.Width := 6.0, [7].Andco_Values.Rate := 4292.5586, [7].Andco_Values.Pounds_Per_Inch := 65.0, [7].Andco_Values.New_Rate := 3700.0, [7].Andco_Values.Analog := 1, [7].Andco_Values.Min_Position := 6, [7].Andco_Values.Length := 12.0, [7].Andco_Values.InchesOpen := 11.575781, [7].Andco_Values.AnalogValue := 9884, [7].Clean_Load_Delay_Stop := 36500, [7].Treat_Load_Delay_Stop := 33000, [7].tmrStopDelay.EN := 1, [7].tmrStopDelay.TT := 1, [7].Available_For_Clean_Load := 1, [7].Available_For_Treat_Load := 1, [8].Bin_Description := '12', [8].Bin_Variety.Name := 'Empty', [8].Bin_Variety.Color[0].Color := 1, [8].Rate_Cal_Points[1].Andco_Position := 3358, [8].Rate_Cal_Points[1].Rate := 1000, [8].Rate_Cal_Points[2].Andco_Position := 5110, [8].Rate_Cal_Points[2].Rate := 2000, [8].Rate_Cal_Points[3].Andco_Position := 6534, [8].Rate_Cal_Points[3].Rate := 3000, [8].Rate_Cal_Points[4].Andco_Position := 8210, [8].Rate_Cal_Points[4].Rate := 4000,
        [8].Clean_Load_Delay_Start := 37000, [8].Treat_Load_Delay_Start := 31000, [8].Andco_Values.Cal_Status := 4, [8].Andco_Values.Raw_Position := 8474, [8].Andco_Values.Max_Position := 15055, [8].Andco_Values.Preact := 20, [8].Andco_Values.Percent_Open := 0.66141117, [8].Andco_Values.New_Pos := 61, [8].Andco_Values.Width := 6.0, [8].Andco_Values.Rate := 4157.518, [8].Andco_Values.Pounds_Per_Inch := 65.0, [8].Andco_Values.New_Rate := 3800.0, [8].Andco_Values.Analog := 1, [8].Andco_Values.Min_Position := 2243, [8].Andco_Values.Length := 12.0, [8].Andco_Values.InchesOpen := 7.936934, [8].Andco_Values.AnalogValue := 10717, [8].Clean_Load_Delay_Stop := 37000, [8].Treat_Load_Delay_Stop := 34000, [8].tmrStopDelay.EN := 1, [8].tmrStopDelay.TT := 1, [8].Available_For_Clean_Load := 1, [8].Available_For_Treat_Load := 1, [9].Bin_Description := '14', [9].Bin_Variety.Item_Number := '873002', [9].Bin_Variety.Name := 'HD-307 CERTIFIED HWW', [9].Bin_Variety.Class := 'Certified', [9].Bin_Variety.Color[0].Color := 1, [9].Rate_Cal_Points[1].Andco_Position := 2158, [9].Rate_Cal_Points[1].Rate := 1000, [9].Rate_Cal_Points[2].Andco_Position := 4887, [9].Rate_Cal_Points[2].Rate := 2000, [9].Rate_Cal_Points[3].Andco_Position := 6612, [9].Rate_Cal_Points[3].Rate := 3000, [9].Rate_Cal_Points[4].Andco_Position := 8287, [9].Rate_Cal_Points[4].Rate := 4000, [9].Clean_Load_Delay_Start := 37500, [9].Treat_Load_Delay_Start := 31000, [9].Andco_Values.Raw_Position := 8668, [9].Andco_Values.Max_Position := 13031, [9].Andco_Values.Preact := 20, [9].Andco_Values.Percent_Open := 0.68679184, [9].Andco_Values.Width := 6.0, [9].Andco_Values.Rate := 4227.463, [9].Andco_Values.Pounds_Per_Inch := 65.0, [9].Andco_Values.Analog := 1, [9].Andco_Values.Min_Position := 410, [9].Andco_Values.Length := 12.0, [9].Andco_Values.InchesOpen := 8.241502, [9].Andco_Values.AnalogValue := 9078, [9].Clean_Load_Delay_Stop := 37500, [9].Treat_Load_Delay_Stop := 34000, [9].tmrStopDelay.EN := 1, [9].tmrStopDelay.TT := 1, [9].Available_For_Clean_Load := 1, [9].Available_For_Treat_Load := 1, [10].Bin_Description := '15', [10].Bin_Variety.Item_Number := '873002', [10].Bin_Variety.Name := 'HD-307 CERTIFIED HWW', [10].Bin_Variety.Class := 'Certified',
        [10].Bin_Variety.Color[0].Color := 1, [10].Rate_Cal_Points[1].Andco_Position := 2321, [10].Rate_Cal_Points[1].Rate := 1000, [10].Rate_Cal_Points[2].Andco_Position := 4523, [10].Rate_Cal_Points[2].Rate := 2000, [10].Rate_Cal_Points[3].Andco_Position := 6483, [10].Rate_Cal_Points[3].Rate := 3000, [10].Rate_Cal_Points[4].Andco_Position := 8309, [10].Rate_Cal_Points[4].Rate := 4000, [10].Clean_Load_Delay_Start := 38000, [10].Treat_Load_Delay_Start := 30000, [10].Andco_Values.Cal_Status := 4, [10].Andco_Values.Raw_Position := 8354, [10].Andco_Values.Max_Position := 12922, [10].Andco_Values.Preact := 20, [10].Andco_Values.Percent_Open := 0.6724082, [10].Andco_Values.Width := 6.0, [10].Andco_Values.Rate := 4024.644, [10].Andco_Values.Pounds_Per_Inch := 65.0, [10].Andco_Values.Analog := 1, [10].Andco_Values.Min_Position := 498, [10].Andco_Values.Length := 12.0, [10].Andco_Values.InchesOpen := 8.068899, [10].Andco_Values.AnalogValue := 8852, [10].Clean_Load_Delay_Stop := 38000, [10].Treat_Load_Delay_Stop := 34000, [10].tmrStartDelay.PRE := 2000, [10].tmrStopDelay.PRE := 2000, [10].tmrStopDelay.EN := 1, [10].tmrStopDelay.TT := 1, [10].StartDelayPre := 2000, [10].StopDelayPre := 2000, [10].Available_For_Clean_Load := 1, [10].Available_For_Treat_Load := 1, [11].Bin_Description := '20', [11].Bin_Variety.Item_Number := '873003', [11].Bin_Variety.Name := 'DAYN CERTIFIED HWW', [11].Bin_Variety.Class := 'Certified', [11].Bin_Variety.Color[0].Color := 1, [11].Rate_Cal_Points[1].Andco_Position := 3830, [11].Rate_Cal_Points[1].Rate := 1000, [11].Rate_Cal_Points[2].Andco_Position := 5231, [11].Rate_Cal_Points[2].Rate := 2000, [11].Rate_Cal_Points[3].Andco_Position := 7521, [11].Rate_Cal_Points[3].Rate := 3000, [11].Rate_Cal_Points[4].Andco_Position := 8755, [11].Rate_Cal_Points[4].Rate := 4000, [11].Clean_Load_Delay_Start := 38000, [11].Treat_Load_Delay_Start := 31000, [11].Andco_Values.Cal_Status := 2, [11].Andco_Values.Raw_Position := 8988, [11].Andco_Values.Max_Position := 12959, [11].Andco_Values.Preact := 32, [11].Andco_Values.Percent_Open := 0.72712564, [11].Andco_Values.New_Pos := 78, [11].Andco_Values.Width := 6.0, [11].Andco_Values.Rate := 4188.817, [11].Andco_Values.Pounds_Per_Inch := 65.0, [11].Andco_Values.New_Rate := 4400.0, [11].Andco_Values.Analog := 1,
        [11].Andco_Values.Min_Position := 598, [11].Andco_Values.Length := 12.0, [11].Andco_Values.InchesOpen := 8.725508, [11].Andco_Values.AnalogValue := 9586, [11].Clean_Load_Delay_Stop := 38000, [11].Treat_Load_Delay_Stop := 35000, [11].tmrStopDelay.EN := 1, [11].tmrStopDelay.TT := 1, [11].Available_For_Clean_Load := 1, [11].Available_For_Treat_Load := 1, [12].Bin_Description := '13', [12].Bin_Variety.Item_Number := '823072', [12].Bin_Variety.Name := 'VOODOO CF CERTIFIED FALL SWH', [12].Bin_Variety.Class := 'Certified', [12].Bin_Variety.Color[0].Color := 1, [12].Rate_Cal_Points[1].Andco_Position := 2243, [12].Rate_Cal_Points[1].Rate := 1000, [12].Rate_Cal_Points[2].Andco_Position := 4281, [12].Rate_Cal_Points[2].Rate := 2000, [12].Rate_Cal_Points[3].Andco_Position := 5779, [12].Rate_Cal_Points[3].Rate := 3000, [12].Rate_Cal_Points[4].Andco_Position := 7567, [12].Rate_Cal_Points[4].Rate := 4000, [12].Clean_Load_Delay_Start := 38500, [12].Treat_Load_Delay_Start := 32000, [12].Andco_Values.Cal_Status := 2, [12].Andco_Values.Raw_Position := 7647, [12].Andco_Values.Max_Position := 12088, [12].Andco_Values.Preact := 20, [12].Andco_Values.Percent_Open := 0.6331346, [12].Andco_Values.New_Pos := 36, [12].Andco_Values.Width := 6.0, [12].Andco_Values.Rate := 4044.7427, [12].Andco_Values.Pounds_Per_Inch := 65.0, [12].Andco_Values.New_Rate := 2500.0, [12].Andco_Values.Analog := 1, [12].Andco_Values.Min_Position := 10, [12].Andco_Values.Length := 12.0, [12].Andco_Values.InchesOpen := 7.5976152, [12].Andco_Values.AnalogValue := 7657, [12].Clean_Load_Delay_Stop := 38500, [12].Treat_Load_Delay_Stop := 36000, [12].tmrStopDelay.EN := 1, [12].tmrStopDelay.TT := 1, [12].Available_For_Clean_Load := 1, [12].Available_For_Treat_Load := 1, [13].Bin_Description := '19', [13].Bin_Variety.Name := 'Empty', [13].Bin_Variety.Color[0].Color := 1, [13].Rate_Cal_Points[1].Andco_Position := 1992, [13].Rate_Cal_Points[1].Rate := 1000, [13].Rate_Cal_Points[2].Andco_Position := 3762, [13].Rate_Cal_Points[2].Rate := 2000, [13].Rate_Cal_Points[3].Andco_Position := 5733, [13].Rate_Cal_Points[3].Rate := 3000, [13].Rate_Cal_Points[4].Andco_Position := 7278, [13].Rate_Cal_Points[4].Rate := 4000, [13].Clean_Load_Delay_Start := 38500, [13].Treat_Load_Delay_Start := 33000, [13].Andco_Values.Cal_Status := 4,
        [13].Andco_Values.Raw_Position := 7215, [13].Andco_Values.Max_Position := 14383, [13].Andco_Values.Preact := 20, [13].Andco_Values.Percent_Open := 0.5766925, [13].Andco_Values.Width := 6.0, [13].Andco_Values.Rate := 3959.2231, [13].Andco_Values.Pounds_Per_Inch := 65.0, [13].Andco_Values.Analog := 1, [13].Andco_Values.Min_Position := 1872, [13].Andco_Values.Length := 12.0, [13].Andco_Values.InchesOpen := 6.92031, [13].Andco_Values.AnalogValue := 9087, [13].Clean_Load_Delay_Stop := 38500, [13].Treat_Load_Delay_Stop := 36000, [13].tmrStopDelay.EN := 1, [13].tmrStopDelay.TT := 1, [13].Available_For_Clean_Load := 1, [13].Available_For_Treat_Load := 1, [14].Bin_Description := '19 SIDE', [14].Bin_Variety.Name := 'Empty', [14].Rate_Cal_Points[1].Andco_Position := 10, [14].Rate_Cal_Points[1].Rate := 1000, [14].Rate_Cal_Points[2].Andco_Position := 20, [14].Rate_Cal_Points[2].Rate := 2000, [14].Rate_Cal_Points[3].Andco_Position := 43, [14].Rate_Cal_Points[3].Rate := 3000, [14].Rate_Cal_Points[4].Andco_Position := 5025, [14].Rate_Cal_Points[4].Rate := 4000, [14].Clean_Load_Delay_Start := 9000, [14].Treat_Load_Delay_Start := 9000, [14].Andco_Values.Raw_Position := 9078, [14].Andco_Values.Max_Position := 120, [14].Andco_Values.Preact := 20, [14].Andco_Values.Percent_Open := 75.65, [14].Andco_Values.Width := 6.0, [14].Andco_Values.Rate := 4813.529, [14].Andco_Values.Pounds_Per_Inch := 65.0, [14].Andco_Values.Analog := 1, [14].Andco_Values.Length := 12.0, [14].Andco_Values.InchesOpen := 907.80005, [14].Andco_Values.AnalogValue := 9078, [14].Clean_Load_Delay_Stop := 9000, [14].Treat_Load_Delay_Stop := 9000, [14].tmrStartDelay.PRE := 4000, [14].tmrStopDelay.PRE := 4000, [14].tmrStopDelay.EN := 1, [14].tmrStopDelay.TT := 1, [14].StartDelayPre := 4000, [14].StopDelayPre := 4000, [14].Available_For_Clean_Load := 1, [14].Available_For_Treat_Load := 1, [15].Bin_Description := '13 SIDE', [15].Bin_Variety.Name := 'Empty', [15].Rate_Cal_Points[1].Andco_Position := 10, [15].Rate_Cal_Points[1].Rate := 1000, [15].Rate_Cal_Points[2].Andco_Position := 20, [15].Rate_Cal_Points[2].Rate := 2000, [15].Rate_Cal_Points[3].Andco_Position := 43, [15].Rate_Cal_Points[3].Rate := 3000, [15].Rate_Cal_Points[4].Andco_Position := 6367,
        [15].Rate_Cal_Points[4].Rate := 4000, [15].Clean_Load_Delay_Start := 9000, [15].Treat_Load_Delay_Start := 9000, [15].Andco_Values.Raw_Position := 8852, [15].Andco_Values.Max_Position := 120, [15].Andco_Values.Preact := 20, [15].Andco_Values.Percent_Open := 73.76667, [15].Andco_Values.Width := 6.0, [15].Andco_Values.Rate := 4392.9473, [15].Andco_Values.Pounds_Per_Inch := 65.0, [15].Andco_Values.Analog := 1, [15].Andco_Values.Length := 12.0, [15].Andco_Values.InchesOpen := 885.2001, [15].Andco_Values.AnalogValue := 8852, [15].Clean_Load_Delay_Stop := 9000, [15].Treat_Load_Delay_Stop := 9000, [15].tmrStopDelay.EN := 1, [15].tmrStopDelay.TT := 1, [15].Available_For_Clean_Load := 1, [15].Available_For_Treat_Load := 1, [16].Bin_Description := '11', [16].Bin_Variety.Item_Number := '823098', [16].Bin_Variety.Name := 'RE-DAG COAXIUM - CERTIFIED', [16].Bin_Variety.Class := 'Certified', [16].Bin_Variety.Color[0].Color := 1, [16].Rate_Cal_Points[1].Andco_Position := 4978, [16].Rate_Cal_Points[1].Rate := 1000, [16].Rate_Cal_Points[2].Andco_Position := 8166, [16].Rate_Cal_Points[2].Rate := 2000, [16].Rate_Cal_Points[3].Andco_Position := 10647, [16].Rate_Cal_Points[3].Rate := 3000, [16].Rate_Cal_Points[4].Andco_Position := 14081, [16].Rate_Cal_Points[4].Rate := 4000, [16].Clean_Load_Delay_Start := 27000, [16].Treat_Load_Delay_Start := 11000, [16].Bindicator_Low := 1, [16].Andco_Values.Cal_Status := 4, [16].Andco_Values.Raw_Position := 13887, [16].Andco_Values.Max_Position := 16180, [16].Andco_Values.Preact := 20, [16].Andco_Values.Percent_Open := 0.9065213, [16].Andco_Values.New_Pos := 101, [16].Andco_Values.Width := 6.0, [16].Andco_Values.Rate := 3943.506, [16].Andco_Values.Pounds_Per_Inch := 65.0, [16].Andco_Values.New_Rate := 4000.0, [16].Andco_Values.Analog := 1, [16].Andco_Values.Min_Position := 861, [16].Andco_Values.Length := 12.0, [16].Andco_Values.InchesOpen := 10.878256, [16].Andco_Values.AnalogValue := 14748, [16].Clean_Load_Delay_Stop := 27000, [16].Treat_Load_Delay_Stop := 12000, [16].tmrStopDelay.EN := 1, [16].tmrStopDelay.TT := 1, [16].Available_For_Clean_Load := 1, [16].Available_For_Treat_Load := 1, [17].Bin_Description := '12', [17].Bin_Variety.Item_Number := '843022', [17].Bin_Variety.Name := 'VENOM CERTIFIED DNS',
        [17].Bin_Variety.Class := 'Certified', [17].Bin_Variety.Color[0].Color := 1, [17].Rate_Cal_Points[1].Andco_Position := 5131, [17].Rate_Cal_Points[1].Rate := 1000, [17].Rate_Cal_Points[2].Andco_Position := 7438, [17].Rate_Cal_Points[2].Rate := 2000, [17].Rate_Cal_Points[3].Andco_Position := 10479, [17].Rate_Cal_Points[3].Rate := 3000, [17].Rate_Cal_Points[4].Andco_Position := 14378, [17].Rate_Cal_Points[4].Rate := 4000, [17].Clean_Load_Delay_Start := 18390, [17].Treat_Load_Delay_Start := 10000, [17].Andco_Values.Fully_Open := 1, [17].Andco_Values.Cal_Status := 4, [17].Andco_Values.Raw_Position := 14945, [17].Andco_Values.Max_Position := 15450, [17].Andco_Values.Preact := 55, [17].Andco_Values.Percent_Open := 0.9995318, [17].Andco_Values.New_Pos := 108, [17].Andco_Values.Width := 6.0, [17].Andco_Values.Rate := 4145.422, [17].Andco_Values.Pounds_Per_Inch := 65.0, [17].Andco_Values.New_Rate := 4000.0, [17].Andco_Values.Analog := 1, [17].Andco_Values.Min_Position := 498, [17].Andco_Values.Length := 12.0, [17].Andco_Values.InchesOpen := 11.994382, [17].Andco_Values.AnalogValue := 15443, [17].Clean_Load_Delay_Stop := 18390, [17].Treat_Load_Delay_Stop := 11000, [17].tmrStopDelay.EN := 1, [17].tmrStopDelay.TT := 1, [17].Available_For_Clean_Load := 1, [17].Available_For_Treat_Load := 1, [18].Bin_Description := '13', [18].Bin_Variety.Name := 'Empty', [18].Bin_Variety.Color[0].Color := 1, [18].Rate_Cal_Points[1].Andco_Position := 4915, [18].Rate_Cal_Points[1].Rate := 1000, [18].Rate_Cal_Points[2].Andco_Position := 7628, [18].Rate_Cal_Points[2].Rate := 2000, [18].Rate_Cal_Points[3].Andco_Position := 12268, [18].Rate_Cal_Points[3].Rate := 3000, [18].Rate_Cal_Points[4].Andco_Position := 13372, [18].Rate_Cal_Points[4].Rate := 4000, [18].Clean_Load_Delay_Start := 17440, [18].Treat_Load_Delay_Start := 10000, [18].Andco_Values.Cal_Status := 2, [18].Andco_Values.Raw_Position := 13995, [18].Andco_Values.Max_Position := 16053, [18].Andco_Values.Preact := 20, [18].Andco_Values.Percent_Open := 0.8855353, [18].Andco_Values.Width := 6.0, [18].Andco_Values.Rate := 4564.3115, [18].Andco_Values.Pounds_Per_Inch := 65.0, [18].Andco_Values.Analog := 1, [18].Andco_Values.Min_Position := 249, [18].Andco_Values.Length := 12.0, [18].Andco_Values.InchesOpen := 10.626424, [18].Andco_Values.AnalogValue := 14244,
        [18].Treat_Load_Delay_Stop := 11000, [18].tmrStopDelay.EN := 1, [18].tmrStopDelay.TT := 1, [18].Available_For_Clean_Load := 1, [18].Available_For_Treat_Load := 1, [19].Bin_Description := '14', [19].Bin_Variety.Item_Number := '822087', [19].Bin_Variety.Name := 'LCS ECLIPSE AX - 0225 COAXIUM REGISTERED HRW', [19].Bin_Variety.Class := 'Registered', [19].Bin_Variety.Color[0].Color := 1, [19].Rate_Cal_Points[1].Andco_Position := 3696, [19].Rate_Cal_Points[1].Rate := 1000, [19].Rate_Cal_Points[2].Andco_Position := 6573, [19].Rate_Cal_Points[2].Rate := 2000, [19].Rate_Cal_Points[3].Andco_Position := 9630, [19].Rate_Cal_Points[3].Rate := 3000, [19].Rate_Cal_Points[4].Andco_Position := 12560, [19].Rate_Cal_Points[4].Rate := 4000, [19].Clean_Load_Delay_Start := 16610, [19].Treat_Load_Delay_Start := 10000, [19].Andco_Values.Cal_Status := 4, [19].Andco_Values.Raw_Position := 12753, [19].Andco_Values.Max_Position := 16151, [19].Andco_Values.Preact := 20, [19].Andco_Values.Percent_Open := 0.8254369, [19].Andco_Values.Width := 6.0, [19].Andco_Values.Rate := 4065.8704, [19].Andco_Values.Pounds_Per_Inch := 65.0, [19].Andco_Values.Analog := 1, [19].Andco_Values.Min_Position := 701, [19].Andco_Values.Length := 12.0, [19].Andco_Values.InchesOpen := 9.905243, [19].Andco_Values.AnalogValue := 13454, [19].Clean_Load_Delay_Stop := 16610, [19].Treat_Load_Delay_Stop := 9000, [19].tmrStopDelay.EN := 1, [19].tmrStopDelay.TT := 1, [19].Available_For_Clean_Load := 1, [19].Available_For_Treat_Load := 1, [20].Bin_Description := '15', [20].Bin_Variety.Item_Number := '803003', [20].Bin_Variety.Name := 'JET CERTIFIED HRW', [20].Bin_Variety.Class := 'Certified', [20].Bin_Variety.Color[0].Color := 1, [20].Rate_Cal_Points[1].Andco_Position := 4509, [20].Rate_Cal_Points[1].Rate := 1000, [20].Rate_Cal_Points[2].Andco_Position := 7812, [20].Rate_Cal_Points[2].Rate := 2000, [20].Rate_Cal_Points[3].Andco_Position := 10414, [20].Rate_Cal_Points[3].Rate := 3000, [20].Rate_Cal_Points[4].Andco_Position := 13301, [20].Rate_Cal_Points[4].Rate := 4000, [20].Clean_Load_Delay_Start := 15870, [20].Treat_Load_Delay_Start := 9000, [20].Andco_Values.Cal_Status := 4, [20].Andco_Values.Raw_Position := 14405, [20].Andco_Values.Max_Position := 15728, [20].Andco_Values.Preact := 20, [20].Andco_Values.Percent_Open := 0.9190965, [20].Andco_Values.New_Pos := 7461,
        [20].Andco_Values.Width := 6.0, [20].Andco_Values.Rate := 4382.404, [20].Andco_Values.Pounds_Per_Inch := 65.0, [20].Andco_Values.New_Rate := 3800.0, [20].Andco_Values.Analog := 1, [20].Andco_Values.Min_Position := 55, [20].Andco_Values.Length := 12.0, [20].Andco_Values.InchesOpen := 11.029159, [20].Andco_Values.AnalogValue := 14460, [20].Treat_Load_Delay_Stop := 9000, [20].tmrStopDelay.EN := 1, [20].tmrStopDelay.TT := 1, [20].Available_For_Clean_Load := 1, [20].Available_For_Treat_Load := 1, [21].Bin_Description := '16', [21].Bin_Variety.Item_Number := '823093', [21].Bin_Variety.Name := 'SCORPION COAX-0291 CERTIFIED SWH', [21].Bin_Variety.Class := 'Certified', [21].Bin_Variety.Color[0].Color := 1, [21].Rate_Cal_Points[1].Andco_Position := 5171, [21].Rate_Cal_Points[1].Rate := 1000, [21].Rate_Cal_Points[2].Andco_Position := 8208, [21].Rate_Cal_Points[2].Rate := 2000, [21].Rate_Cal_Points[3].Andco_Position := 11698, [21].Rate_Cal_Points[3].Rate := 3000, [21].Rate_Cal_Points[4].Andco_Position := 14346, [21].Rate_Cal_Points[4].Rate := 4000, [21].Clean_Load_Delay_Start := 19000, [21].Treat_Load_Delay_Start := 8000, [21].Bindicator_Low := 1, [21].Andco_Values.Cal_Status := 4, [21].Andco_Values.Raw_Position := 5924, [21].Andco_Values.Max_Position := 16315, [21].Andco_Values.Preact := 20, [21].Andco_Values.Percent_Open := 0.37267238, [21].Andco_Values.New_Pos := 133, [21].Andco_Values.Width := 6.0, [21].Andco_Values.Rate := 1247.942, [21].Andco_Values.Pounds_Per_Inch := 65.0, [21].Andco_Values.New_Rate := 5000.0, [21].Andco_Values.Analog := 1, [21].Andco_Values.Min_Position := 419, [21].Andco_Values.Length := 12.0, [21].Andco_Values.InchesOpen := 4.472069, [21].Andco_Values.AnalogValue := 6343, [21].Clean_Load_Delay_Stop := 19000, [21].Treat_Load_Delay_Stop := 9000, [21].tmrStartDelay.PRE := 21000, [21].tmrStopDelay.PRE := 23000, [21].tmrStopDelay.EN := 1, [21].tmrStopDelay.TT := 1, [21].StartDelayPre := 21000, [21].StopDelayPre := 23000, [21].Available_For_Clean_Load := 1, [21].Available_For_Treat_Load := 1, [22].Bin_Description := '17', [22].Bin_Variety.Item_Number := '843036', [22].Bin_Variety.Name := 'HALE CERTIFIED DNS', [22].Bin_Variety.Class := 'Certified', [22].Bin_Variety.Color[0].Color := 1,
        [22].Rate_Cal_Points[1].Andco_Position := 1803, [22].Rate_Cal_Points[1].Rate := 1000, [22].Rate_Cal_Points[2].Andco_Position := 3716, [22].Rate_Cal_Points[2].Rate := 2000, [22].Rate_Cal_Points[3].Andco_Position := 5315, [22].Rate_Cal_Points[3].Rate := 3000, [22].Rate_Cal_Points[4].Andco_Position := 7606, [22].Rate_Cal_Points[4].Rate := 4000, [22].Clean_Load_Delay_Start := 19000, [22].Treat_Load_Delay_Start := 7000, [22].Bindicator_Low := 1, [22].Andco_Values.Cal_Status := 4, [22].Andco_Values.Raw_Position := 7779, [22].Andco_Values.Max_Position := 15450, [22].Andco_Values.Preact := 20, [22].Andco_Values.Percent_Open := 0.5375579, [22].Andco_Values.New_Pos := 47, [22].Andco_Values.Width := 6.0, [22].Andco_Values.Rate := 4075.513, [22].Andco_Values.Pounds_Per_Inch := 65.0, [22].Andco_Values.New_Rate := 4000.0, [22].Andco_Values.Analog := 1, [22].Andco_Values.Min_Position := 979, [22].Andco_Values.Length := 12.0, [22].Andco_Values.InchesOpen := 6.450695, [22].Andco_Values.AnalogValue := 8758, [22].Clean_Load_Delay_Stop := 19000, [22].Treat_Load_Delay_Stop := 10000, [22].tmrStartDelay.PRE := 23000, [22].tmrStopDelay.PRE := 23000, [22].tmrStopDelay.EN := 1, [22].tmrStopDelay.TT := 1, [22].StartDelayPre := 23000, [22].StopDelayPre := 23000, [22].Available_For_Clean_Load := 1, [22].Available_For_Treat_Load := 1, [23].Bin_Description := '21', [23].Bin_Variety.Item_Number := '843001', [23].Bin_Variety.Name := 'BUCK PRONTO CERTIFIED DNS', [23].Bin_Variety.Class := 'Certified', [23].Bin_Variety.Color[0].Color := 1, [23].Rate_Cal_Points[1].Andco_Position := 5036, [23].Rate_Cal_Points[1].Rate := 1000, [23].Rate_Cal_Points[2].Andco_Position := 8241, [23].Rate_Cal_Points[2].Rate := 2000, [23].Rate_Cal_Points[3].Andco_Position := 12245, [23].Rate_Cal_Points[3].Rate := 3000, [23].Rate_Cal_Points[4].Andco_Position := 14788, [23].Rate_Cal_Points[4].Rate := 4000, [23].Clean_Load_Delay_Start := 19000, [23].Treat_Load_Delay_Start := 11000, [23].Bindicator_Low := 1, [23].Andco_Values.Cal_Status := 4, [23].Andco_Values.Raw_Position := 15207, [23].Andco_Values.Max_Position := 16384, [23].Andco_Values.Preact := 20, [23].Andco_Values.Percent_Open := 0.9718796, [23].Andco_Values.New_Pos := 86, [23].Andco_Values.Width := 6.0, [23].Andco_Values.Rate := 4164.766,
        [23].Andco_Values.Pounds_Per_Inch := 65.0, [23].Andco_Values.New_Rate := 4000.0, [23].Andco_Values.Analog := 1, [23].Andco_Values.Min_Position := 737, [23].Andco_Values.Length := 12.0, [23].Andco_Values.InchesOpen := 11.662556, [23].Andco_Values.AnalogValue := 15944, [23].Clean_Load_Delay_Stop := 19000, [23].Treat_Load_Delay_Stop := 14000, [23].tmrStopDelay.EN := 1, [23].tmrStopDelay.TT := 1, [23].Available_For_Clean_Load := 1, [23].Available_For_Treat_Load := 1, [24].Bin_Description := '22', [24].Bin_Variety.Item_Number := '843002', [24].Bin_Variety.Name := 'EXPRESSO CERTIFIED DNS', [24].Bin_Variety.Class := 'Certified', [24].Bin_Variety.Color[0].Color := 1, [24].Rate_Cal_Points[1].Andco_Position := 5147, [24].Rate_Cal_Points[1].Rate := 1000, [24].Rate_Cal_Points[2].Andco_Position := 8427, [24].Rate_Cal_Points[2].Rate := 2000, [24].Rate_Cal_Points[3].Andco_Position := 12356, [24].Rate_Cal_Points[3].Rate := 3000, [24].Rate_Cal_Points[4].Andco_Position := 14863, [24].Rate_Cal_Points[4].Rate := 4000, [24].Clean_Load_Delay_Start := 23500, [24].Treat_Load_Delay_Start := 14000, [24].Bindicator_Low := 1, [24].Andco_Values.Cal_Status := 4, [24].Andco_Values.Raw_Position := 14817, [24].Andco_Values.Max_Position := 16384, [24].Andco_Values.Preact := 20, [24].Andco_Values.Percent_Open := 0.9250796, [24].Andco_Values.New_Pos := 57, [24].Andco_Values.Width := 6.0, [24].Andco_Values.Rate := 3981.6514, [24].Andco_Values.Pounds_Per_Inch := 65.0, [24].Andco_Values.New_Rate := 2000.0, [24].Andco_Values.Analog := 1, [24].Andco_Values.Min_Position := 367, [24].Andco_Values.Length := 12.0, [24].Andco_Values.InchesOpen := 11.100955, [24].Andco_Values.AnalogValue := 15184, [24].Clean_Load_Delay_Stop := 23500, [24].Treat_Load_Delay_Stop := 15000, [24].tmrStartDelay.PRE := 15000, [24].tmrStopDelay.PRE := 17000, [24].tmrStopDelay.EN := 1, [24].tmrStopDelay.TT := 1, [24].StartDelayPre := 15000, [24].StopDelayPre := 17000, [24].Available_For_Clean_Load := 1, [24].Available_For_Treat_Load := 1, [25].Bin_Description := '23', [25].Bin_Variety.Item_Number := '843022', [25].Bin_Variety.Name := 'VENOM CERTIFIED DNS', [25].Bin_Variety.Class := 'Certified', [25].Rate_Cal_Points[1].Andco_Position := 4846, [25].Rate_Cal_Points[1].Rate := 1000,
        [25].Rate_Cal_Points[2].Andco_Position := 8120, [25].Rate_Cal_Points[2].Rate := 2000, [25].Rate_Cal_Points[3].Andco_Position := 11636, [25].Rate_Cal_Points[3].Rate := 3000, [25].Rate_Cal_Points[4].Andco_Position := 13864, [25].Rate_Cal_Points[4].Rate := 4000, [25].Clean_Load_Delay_Start := 28000, [25].Treat_Load_Delay_Start := 18000, [25].Bindicator_Low := 1, [25].Andco_Values.Cal_Status := 4, [25].Andco_Values.Raw_Position := 14906, [25].Andco_Values.Max_Position := 16033, [25].Andco_Values.Preact := 20, [25].Andco_Values.Percent_Open := 0.9807869, [25].Andco_Values.New_Pos := 8762, [25].Andco_Values.Width := 6.0, [25].Andco_Values.Rate := 4467.684, [25].Andco_Values.Pounds_Per_Inch := 65.0, [25].Andco_Values.New_Rate := 3800.0, [25].Andco_Values.Analog := 1, [25].Andco_Values.Min_Position := 835, [25].Andco_Values.Length := 12.0, [25].Andco_Values.InchesOpen := 11.7694435, [25].Andco_Values.AnalogValue := 15741, [25].Clean_Load_Delay_Stop := 28000, [25].Treat_Load_Delay_Stop := 20000, [25].tmrStopDelay.EN := 1, [25].tmrStopDelay.TT := 1, [25].Available_For_Clean_Load := 1, [25].Available_For_Treat_Load := 1, [26].Bin_Description := '24', [26].Bin_Variety.Item_Number := '803003', [26].Bin_Variety.Name := 'JET CERTIFIED HRW', [26].Bin_Variety.Class := 'Certified', [26].Bin_Variety.Color[0].Color := 1, [26].Rate_Cal_Points[1].Andco_Position := 5096, [26].Rate_Cal_Points[1].Rate := 1000, [26].Rate_Cal_Points[2].Andco_Position := 8425, [26].Rate_Cal_Points[2].Rate := 2000, [26].Rate_Cal_Points[3].Andco_Position := 12377, [26].Rate_Cal_Points[3].Rate := 3000, [26].Rate_Cal_Points[4].Andco_Position := 14785, [26].Rate_Cal_Points[4].Rate := 4000, [26].Clean_Load_Delay_Start := 23000, [26].Treat_Load_Delay_Start := 16000, [26].Andco_Values.Cal_Status := 4, [26].Andco_Values.Raw_Position := 14844, [26].Andco_Values.Max_Position := 16384, [26].Andco_Values.Preact := 20, [26].Andco_Values.Percent_Open := 0.93071663, [26].Andco_Values.New_Pos := 76, [26].Andco_Values.Width := 6.0, [26].Andco_Values.Rate := 4024.5017, [26].Andco_Values.Pounds_Per_Inch := 65.0, [26].Andco_Values.New_Rate := 3800.0, [26].Andco_Values.Analog := 1, [26].Andco_Values.Min_Position := 435, [26].Andco_Values.Length := 12.0, [26].Andco_Values.InchesOpen := 11.1686, [26].Andco_Values.AnalogValue := 15279,
        [26].Clean_Load_Delay_Stop := 23000, [26].Treat_Load_Delay_Stop := 16000, [26].tmrStartDelay.PRE := 5000, [26].tmrStopDelay.PRE := 8000, [26].tmrStopDelay.EN := 1, [26].tmrStopDelay.TT := 1, [26].StartDelayPre := 5000, [26].StopDelayPre := 8000, [26].Available_For_Clean_Load := 1, [26].Available_For_Treat_Load := 1, [27].Bin_Description := '25', [27].Bin_Variety.Item_Number := '823087', [27].Bin_Variety.Name := 'LCS ECLIPSE AX - 0225 COAXIUM CERTIFIED HRW', [27].Bin_Variety.Class := 'Certified', [27].Bin_Variety.Color[0].Color := 1, [27].Rate_Cal_Points[1].Andco_Position := 5099, [27].Rate_Cal_Points[1].Rate := 1000, [27].Rate_Cal_Points[2].Andco_Position := 8615, [27].Rate_Cal_Points[2].Rate := 2000, [27].Rate_Cal_Points[3].Andco_Position := 12478, [27].Rate_Cal_Points[3].Rate := 3000, [27].Rate_Cal_Points[4].Andco_Position := 14424, [27].Rate_Cal_Points[4].Rate := 4000, [27].Clean_Load_Delay_Start := 27000, [27].Treat_Load_Delay_Start := 17000, [27].Bindicator_Low := 1, [27].Andco_Values.Cal_Status := 4, [27].Andco_Values.Raw_Position := 14595, [27].Andco_Values.Max_Position := 16121, [27].Andco_Values.Preact := 20, [27].Andco_Values.Percent_Open := 0.9062403, [27].Andco_Values.Width := 6.0, [27].Andco_Values.Rate := 4087.8726, [27].Andco_Values.Pounds_Per_Inch := 65.0, [27].Andco_Values.Analog := 1, [27].Andco_Values.Min_Position := 16, [27].Andco_Values.Length := 12.0, [27].Andco_Values.InchesOpen := 10.874884, [27].Andco_Values.AnalogValue := 14611, [27].Clean_Load_Delay_Stop := 27000, [27].Treat_Load_Delay_Stop := 21000, [27].tmrStopDelay.EN := 1, [27].tmrStopDelay.TT := 1, [27].Available_For_Clean_Load := 1, [27].Available_For_Treat_Load := 1, [28].Bin_Description := '26', [28].Bin_Variety.Item_Number := '803021', [28].Bin_Variety.Name := 'LCS BLACKBIRD CERTIFIED HRW', [28].Bin_Variety.Class := 'Certified', [28].Bin_Variety.Color[0].Color := 1, [28].Rate_Cal_Points[1].Andco_Position := 3558, [28].Rate_Cal_Points[1].Rate := 1000, [28].Rate_Cal_Points[2].Andco_Position := 7029, [28].Rate_Cal_Points[2].Rate := 2000, [28].Rate_Cal_Points[3].Andco_Position := 10092, [28].Rate_Cal_Points[3].Rate := 3000, [28].Rate_Cal_Points[4].Andco_Position := 13120, [28].Rate_Cal_Points[4].Rate := 4000, [28].Clean_Load_Delay_Start := 31000, [28].Treat_Load_Delay_Start := 21000,
        [28].Bindicator_Low := 1, [28].Andco_Values.Cal_Status := 4, [28].Andco_Values.Raw_Position := 15129, [28].Andco_Values.Max_Position := 15233, [28].Andco_Values.Preact := 20, [28].Andco_Values.Percent_Open := 0.994217, [28].Andco_Values.New_Pos := 95, [28].Andco_Values.Width := 6.0, [28].Andco_Values.Rate := 4663.474, [28].Andco_Values.Pounds_Per_Inch := 65.0, [28].Andco_Values.New_Rate := 3800.0, [28].Andco_Values.Analog := 1, [28].Andco_Values.Min_Position := 16, [28].Andco_Values.Length := 12.0, [28].Andco_Values.InchesOpen := 11.930604, [28].Andco_Values.AnalogValue := 15145, [28].Clean_Load_Delay_Stop := 31000, [28].Treat_Load_Delay_Stop := 24000, [28].tmrStopDelay.EN := 1, [28].tmrStopDelay.TT := 1, [28].Available_For_Clean_Load := 1, [28].Available_For_Treat_Load := 1);
   Loadout_K_Valve : udt_Loadout_K_Valve[2] := ([0].Clean_Gate_Opened := 1, [1].Clean_Gate_Opened := 1);
   Loadout_K_Valve_Control : Loadout_K_Valve_Control[2];
   Loadout_KValve_Not_Used : BOOL;
   Longest_Clean_IDX : DINT := 21;
   Longest_Clean_Start_IDX : DINT;
   Longest_Clean_Start_Time : DINT;
   Longest_Clean_Stop_IDX : DINT;
   Longest_Clean_Stop_Time : DINT;
   Longest_Clean_Time : DINT;
   Longest_IDX : DINT := 5;
   Longest_Time : DINT := 60000;
   Longest_Time_IDX : DINT;
   Longest_Treat_IDX : DINT;
   Longest_Treat_Start_IDX : DINT;
   Longest_Treat_Start_Time : DINT;
   Longest_Treat_Stop_IDX : DINT;
   Longest_Treat_Stop_Time : DINT;
   Longest_Treat_Time : DINT;
   Loop_Idx : DINT := 14;
   Man_Start_Stop_Allowed : BOOL := 1;
   Manual_Blow_Out : BOOL;
   Manual_Mode : BOOL;
   Manual_Open_Calibration_Valves : BOOL;
   Manually_Start_Treater : BOOL;
   Move_Bin_Config : BOOL;
   NA : BOOL;
   New_DeltaX : REAL := -23.0;
   New_DeltaY : REAL := -1000.0;
   Ok_Stop_Belt : BOOL;
   Open_Clean_Bins : BOOL;
   Open_Transfer_Bins : BOOL;
   Open_Treat_Bins : BOOL;
   Pause_Load : BOOL;
   Pause_Load_By_Time : BOOL[32];
   Pause_Load_By_Weight : BOOL[32];
   Pause_Load_Expired : DINT[2];
   Pause_Load_Pre : DINT[2] := ([0] := 29000, [1] := 32000);
   Pause_Transfer_By_Time : BOOL;
   Pause_Transfer_Load_Expired : DINT;
   Pause_Transfer_Msc : DINT := 1800000;
   Pause_Transfer_Pre : DINT := 30;
   Pause_Treat_By_Time : BOOL;
   Pause_Treat_Pre : DINT;
   Pause_Treatment : BOOL;
   Point1 : DINT := 3;
   Point2 : DINT := 4;
   Probe_Above_K_Valve : BOOL;
   Produced_Motor_Values : DINT;
   Rate_Mult : REAL := 0.33025098;
   Remote_Pause_Treat : BOOL;
   Request_Variety : udt_Requested_Variety := (Item_Number := '123', Percentage := 1.0, Bin_Available := 1);
   Requested_Varieties : udt_Requested_Variety[10] := ([0].Item_Number := '123456', [0].Percentage := 0.5, [0].Bin_Available := 1);
   Reset_Bin_Cal : BOOL := 1;
   Reset_Remote_Pause : BOOL;
   Reset_Treat_Chemicals : BOOL;
   ResetSelectedBins : BOOL := 1;
   Rev_Delay_Latch_FWD : BOOL;
   Rev_Delay_Latch_REV : BOOL;
   Reverse_Belt_Forward_Interlock : BOOL := 1;
   Reverse_Belt_Stopping : BOOL;
   Reversing_Belt_Bypass_Valve : BOOL := 1;
   Reversing_Belt_Fans : udt_Cyclone;
   Reversing_Belt_Name : STRING; {constant}
   Reversing_Belt_Reversed : BOOL;
   Scale : SCALE;
   Scale_Target : DINT;
   SCL_01 : SCALE;
   SCL_02 : SCALE;
   SCL_03 : SCALE;
   SCL_04 : SCALE;
   SCL_05 : SCALE;
   SCL_06 : SCALE;
   SCL_07 : SCALE;
   SCL_08 : SCALE := (InRawMax := 30000.0, InEUMax := 50.0);
   SCL_16 : SCALE := (In := 3976.0, InRawMax := 20000.0, InRawMin := 4000.0, InEUMax := 200.0, Out := -0.3, MinAlarm := 1);
   SCL_AMP_Belt10 : SCALE := (In := 10.0, InRawMax := 30151.0, InEUMax := 50.0, Out := 0.016583197);
   SCL_AMP_Belt11 : SCALE := (In := -1.0, InRawMax := 30154.0, InEUMax := 50.0, Out := -0.0016581548, MinAlarm := 1);
   SCL_AMP_Belt11_01 : SCALE;
   SCL_AMP_Belt7 : SCALE := (In := -53.0, InRawMax := 41874.0, InEUMax := 200.0, Out := -0.2531404, MinAlarm := 1);
   SCL_AMP_Belt7_01 : SCALE;
   SCL_AMP_Belt8 : SCALE := (In := 1.0, InRawMax := 29984.0, InEUMax := 50.0, Out := 0.001667556);
   SCL_AMP_Belt8_01 : SCALE;
   SCL_AMP_Belt9 : SCALE := (In := 18.0, InRawMax := 30000.0, InEUMax := 50.0, Out := 0.030000001);
   SCL_AMP_BIN16_AUG : SCALE := (InRawMax := 30000.0, InEUMax := 50.0);
   SCL_AMP_Bin17_AUG : SCALE;
   SCL_AMPS_Belt4 : SCALE := (In := -11.0, InRawMax := 41623.0, InEUMax := 200.0, Out := -0.05285539, MinAlarm := 1);
   SCL_AMPS_Belt5 : SCALE := (In := 11.0, InRawMax := 30168.0, InEUMax := 50.0, Out := 0.018231237);
   SCL_AMPS_Belt6 : SCALE := (In := 8.0, InRawMax := 30203.0, InEUMax := 50.0, Out := 0.013243717);
   Select_Bin_Load_Type : DINT;
   Select_Bin_To_Cal : BOOL;
   Slope : REAL := 1.992;
   Sort_Time_Idx : DINT;
   Sorted_Times : DINT[29,2];
   Start_Bin_Cal : BOOL;
   Start_Blower_707 : BOOL;
   Start_Clean_Belts_Enabled : BOOL;
   Start_Rev_Mtr : udt_Motor_Start;
   Start_Treat_Belts_Enabled : BOOL;
   Steel_Bin_Timing_Offset : DINT := -5;
   Steel_Rqd_Belts_Running : BOOL;
   Stop_Treater : BOOL;
   SUBTest1 : DINT;
   SubTest2 : DINT;
   System_In_Use : BOOL;
   System_Status_Msg : STRING := 'System$0D$0AIdle';
   System_Status_Msgs : STRING[20] := ([0] := 'System$0D$0AIdle', [1] := 'Manual Mode$0D$0A NO INTERLOCKS ! $0D$0A (Be Careful)');
   Target_Weight : DINT[2] := ([0] := 18800, [1] := 78000);
   Test1 : BOOL;
   Test_10Slp : BOOL;
   Test_20Slp : BOOL := 1;
   Test_Air_Gate : BOOL;
   Test_Air_Gate25 : BOOL;
   Test_Air_Open_Input : BOOL;
   Test_In : BOOL;
   Test_Int : DINT;
   Test_Plug : BOOL;
   TestAmps : DINT;
   TestReal : REAL := 1.235;
   Time_Sorter : CONTROL := (LEN := 29);
   Timed_Gate_Met : DINT;
   Timer_Target : REAL;
   tmr_Auto_Start : TIMER := (PRE := 1000, ACC := 1005);
   tmr_Blow_Out : TIMER := (ACC := 16, EN := 1, DN := 1);
   TMR_Concrete_Fan : TIMER := (PRE := 180000, ACC := 180014);
   TMR_Max_Clean_Delay : TIMER;
   TMR_Max_Treat_Delay : TIMER;
   tmr_Pause_Load_Timer : TIMER[2] := ([0].PRE := 29000, [1].PRE := 32000);
   tmr_Pause_Transfer_Timer : TIMER := (PRE := 1800000);
   tmr_Pause_Treat_Timer : TIMER;
   TMR_Reverse_Delay : TIMER := (PRE := 4000, ACC := 4001);
   tmr_Setpoint : TIMER;
   tmrBin_Delay_Start : TIMER[30] := ([0].PRE := 10000, [0].ACC := 10008, [0].EN := 1, [0].DN := 1, [1].PRE := 5000);
   tmrCleanSetpoint : TIMER;
   tmrCleanTime : TIMER := (PRE := 1000);
   tmrDelayTreatStart : TIMER := (PRE := 30000);
   tmrDelayTreatStop : TIMER := (PRE := 33000);
   tmrResetChemicals : TIMER := (PRE := 1000);
   tmrTransferTime : TIMER := (PRE := 1000);
   tmrTreatSetpoint : TIMER;
   tmrTreatTime : TIMER := (PRE := 1000);
   Transfer_Batch_Status : DINT;
   Transfer_Belts_Starting : BOOL;
   Transfer_From_IDX : DINT := -1;
   Transfer_Interlock : BOOL;
   Transfer_To_IDX : DINT := -1;
   TransferHours : DINT;
   TransferMinuets : DINT;
   TransferSeconds : DINT;
   Treat_Batch_Status : DINT;
   Treat_Bin_Gates_Opened : BOOL := 1;
   Treat_Bins_Open : BOOL;
   Treat_Bins_Ready : BOOL := 1;
   Treat_Interlock : BOOL;
   Treat_Jump_Interlock : BOOL;
   Treat_Load : BOOL;
   Treat_Scale_Target : DINT;
   Treat_Scale_Unavailable : BOOL;
   Treater_Calibration : BOOL;
   Treater_Loadout : udt_Treater_Loadout := (Use_A_Treater := 1, Use_B_Treater := 1, Drip_Gate_Closed := 1);
   Treater_Loadout_Open_Bins : BOOL;
   TreatHours : DINT;
   Treatment_Running : BOOL;
   Treatment_Started : BOOL;
   TreatMinuets : DINT;
   TreatSeconds : DINT;
   Truck_Scale_Control : Truck_Scale_Control[3];
   Use_Concrete_Side_Clean : BOOL;
   Use_Concrete_Side_Treat : BOOL;
   Use_Steel_Side_Clean : BOOL;
   Use_Steel_Side_Treat : BOOL;
   Use_Steel_Transfer_Bins : BOOL;
   X1 : REAL;
   X2 : REAL := 1000.0;
   Y1 : REAL;
   Y2 : REAL := 1992.0;
   ZZTEST : udt_Motor_Start;
END_VAR
